(* IEC 61131-3 sources: SortJet_MasterSPS_Aufbau.fbsproj/11_MMI_Kommunikation, 12 files *)

(* ---- MMI_CONST.gvl ---- *)
(* METADATA
{
	"v3Meta": {
		"objectGuid": "b42c2871-ef06-40a1-9ac4-06faa3b26b72"
	}
}
*)
{attribute 'allow_unqualified_access'}
NAMESPACE MMI_CONST
VAR_GLOBAL CONSTANT

  sSpsVersion                                      : STRING(25) := 'ISO Sortierung V4.0.0.0';

// ************************ START SPS Nachrichtennummern *****************

  SB0_SPS_SPSVERSION                                 : WORD := 32768;
  SB0_SPS_MSG_ERROR                                  : WORD := 32767;
  SB0_SPS_ERROR                                      : WORD := 32766;
  SB0_SPS_WARNUNG                                    : WORD := 32765;
  SB0_SPS_HINWEIS                                    : WORD := 32764;
  SB0_SPS_PARAMETER_CRC                              : WORD := 32763;
  SB0_SPS_DEBUG                                      : WORD := 32762;
  SB0_SPS_DEBUG_TRACE                                : WORD := 32761; // Nachricht die in ein seperates Log-File geschrieben wird ( Void- Message )
  SB0_SPS_LOGSTRING                                  : WORD := 32770; // Nachricht um einen String (60 Zeichen) in das Log zu schreiben

// Nachricht von der SPS zum MMI
  SB0_SPS_SETBETRIEBSART                             : WORD :=  1;
  SB0_SPS_SORTIERUNGQUITTINPUTINQUEUE                : WORD :=  2;
  SB0_SPS_SORTIERUNGQUITTUNGVONISOLINIE              : WORD := 11;
  SB0_SPS_SORTIERUNGQUITTEXTRACTIONSHUTTLEDATA       : WORD := 13;
  SB0_SPS_SORTIERUNGRACKINPOS                        : WORD := 19;
  SB0_SPS_SORTIERUNGRACKSTATIONSTATUS                : WORD := 23;
  SB0_SPS_ERRORMSG                                   : WORD := 30;
  SB0_SPS_TRANSPORTSTATE                             : WORD := 35; // Antwort auf Eckübergabenstatus 0 = Rücktransport / 1 = Weitertransoport
  SB0_SPS_RACKONLOADINGSTATION                       : WORD := 37; // Fächerwagen auf Füllstation angedockt
  SB0_SPS_RACKLOGIN                                  : WORD := 38; // Fächerwagen auf Einschleusestation angedockt
  SB0_SPS_STATUSRACKSTATION                          : WORD := 39; // Antwort auf die Nachricht: SB0_SPS_STATUSRACKSTATION
  SB0_SPS_SETSTATUSLOADINGSTATIONS                   : WORD := 44; // Antwort auf REQUESTSTATUSLOADINGSTATIONS mit 1 = frei; 2 = belegt; 0 = ungültig
  SB0_SPS_SHEETREMOVEDAPPROVALWALL                   : WORD := 45;
  SB0_SPS_SHEETONINPUTTABLE                          : WORD := 46;
  SB0_SPS_RACKPOSITION                               : WORD := 48;
  SB0_SPS_TURNSTATIONPOSITION                        : WORD := 49;

  SB0_SPS_SYSTEMCHECKFINISHED                        : WORD := 51;
  SB0_SPS_SETSHEETSONSHUTTLE                         : WORD := 53;
  SB0_SPS_STATIONSTATUS                              : WORD := 62;
  SBO_SPS_STATIONSEVENT                              : word := 65;
  SB0_SPS_GETSTATIONSTATUS                           : WORD := 67; // BEKOMMEN: Einen Station-Status bekommen -> SystemCheck: Ein/ Austransport etc.
  SB0_SPS_SETSHEETSONSTATION                         : WORD := 68; // Nachricht an die Oberflaeche fuer die Glasmessung auf den Stationen
  SB0_SPS_SORTIERUNGSHUTTLEPOS                       : WORD := 69;
  SB0_SPS_SHUTTLEVORABPOSITIONIERUNGUPDATE           : WORD := 70;
  SB0_SPS_QUITTSHUTTLEVORABPOSITIONIERUNG            : WORD := 71;
  SB0_SPS_SHUTTLEVORABPOSITIONIERUNGABBRUCH          : WORD := 72;
  SB0_SPS_SHUTTLEVORABPOSITIONIERUNGREADY            : WORD := 73;
  SB0_SPS_TRANSFERSHUTTLEFEHLER                      : WORD := 75;
  SB0_SPS_FACHAUFNAHMEDATEN                          : WORD := 76;
  SB0_SPS_TRANSFERSHUTTLECHECK_ABGESCHLOSSEN         : WORD := 77;
  SB0_SPS_LIFTEDTRANSFERSHUTTLEPOSITION              : WORD := 78;
  SB0_SPS_SCHNITTSTELLENDATENFREMDANLAGE             : WORD := 79;

  SB0_SPS_POSITIONMEASUREDATA                        : WORD := 81; // Fächerwagensuche: Wort 0 = (int) SPS Nr Shuttle  / Wort 1+2 = (real) Position rechte (?) Kante der Folie[-1 für nicht gefunden]
  SB0_SPS_HANDFUNKTION_STATUS                        : WORD := 82; // Antwort auf SB0_MMI_SETHANDFUNKTION [22]
  SB0_SPS_SHUTTLEHANDFUNKTION_STATUS                 : WORD := 83; // Antwort auf SB0_MMI_SETSHUTTLEHANDFUNKTION [23]
  SB0_SPS_WATCHDOGTEST                               : WORD := 99;
  SB0_SPS_TRANSFERSHUTTLEBUFFERSLOTPOS               : WORD := 100;
  SB0_SPS_QUIT_SHEET_ORDER                           : WORD := 101;
  SB0_SPS_QUIT_CARRIER_POSITION                      : WORD := 102;
  SB0_SPS_STATION_UPDATE                             : WORD := 110;

// ************************ START MMI Nachrichtennummern *****************
  SB0_MMI_SPSVERSION                                 : WORD := 32768;
  SB0_MMI_GETBETRIEBSART                             : WORD :=  1;
  SB0_MMI_SORTIERUNGINPUTINQUEUE                     : WORD :=  2;
  SB0_MMI_SORTIERUNGCHECKINPUTQUEUE                  : WORD :=  5;
  SB0_MMI_SORTIERUNGCANCELQUEUEDATA                  : WORD :=  7;
  SB0_MMI_SORTIERUNGCANCELISOLINEEVENT               : WORD :=  8; // ISO- Line Event stoppen [Cancel]
  SB0_MMI_SORTIERUNGCANCELSHUTTLEDATA                : WORD :=  9;
  SB0_MMI_SORTIERUNGFAECHERWAGENBALDVOLL             : WORD := 10; // Faecherwagen in der Station bald voll
  SB0_MMI_SORTIERUNGAUTOMATIKSTART                   : WORD := 11;
  SB0_MMI_SORTIERUNGAUTOMATIK_STOP                   : WORD := 12;
  SB0_MMI_SORTIERUNGINSERTEXTRACTIONSHUTTLEDATA      : WORD := 14;
  SB0_MMI_SORTIERUNGFAECHERWAGENWECHSEL              : WORD := 15;
  SB0_MMI_SETHANDFUNKTION                            : WORD := 22;
  SB0_MMI_SETSHUTTLEHANDFUNKTION                     : WORD := 23;
  SB0_MMI_MEASSURERESULT                             : WORD := 30; // Scheibenmessung OK -> Freigabe für die Eckübergabe des Sortjets  0 = nicht OK / 1 = OK
  SB0_MMI_ISOQUITTUNG                                : WORD := 31; // unabhängige Quittung der Sondergläser durch Tasterdruck anfordern
  SB0_MMI_RELEASERACKLOGIN                           : WORD := 39; // Freigabe, dass der Fächerwagen eingeschleußt werden darf
  SB0_MMI_GETSTATUSRACKSTATION                       : WORD := 40; // Anfrage vom MMI nach dem Status einer EINZELNEN Fächerwagenstation => belegt, Muting OK, RFID-Nr.
  SB0_MMI_DOCKRACK                                   : WORD := 41; // Freigabe den AGV Fächerwagen einzuschleusen bzw. das Tor zu öffnen  /  release to open the door for the AGV harp rack
  SB0_MMI_REQUESTSTATUSLOADINGSTATIONS               : WORD := 43; // Anfrage der Oberfläche welche Fächerwagenbeladestationen belegt sind
  SB0_MMI_SETSLOTSFORSHUTTLECHECK                    : WORD := 44; // Anfrage der aktuellen Shuttlepositionnen für den bevorstehenden Check der Maschine
  SB0_MMI_REQUESTTILTSTATION                         : WORD := 51;
  SB0_MMI_SHUTTLEVORABPOSITIONIERUNG                 : WORD := 53; // Shuttle Vorapositionieren falls ein Transfershuttle (welches benötigt wird) gerade beschäftigt ist
  SB0_MMI_FACHAUFNAHMESTART                          : WORD := 55;
  SB0_MMI_POSITIONMEASUREONOFF                       : WORD := 56; // FächerwagenSUCHE    Wort 0 = (int) 1 für AN oder 0 für AUS / Wort 2 = (int) SPS Nr Shuttle
  SB0_MMI_STATIONSTATUS                              : WORD := 67; // Stationsstatus [Antwort in welchem Modus sich die Station befunden hat -> SystemCheck]
  SB0_MMI_SYSTEMCHECKSTATION                         : WORD := 68; // Stationsstatus [Antwort in welchem Modus sich die Station befunden hat -> SystemCheck]
  SB0_MMI_GETSORTIERUNGSHUTTLEPOS                    : WORD := 69;
  SB0_MMI_IOANZEIGE_AKTIVIEREN_DEAKTIVIEREN          : WORD := 70; // Anzeige der IO´s im MMI Service  WORT 0: 1 = sichtbar / 0 = unsichtbar
  SB0_MMI_AUFTRAGSDATEN_FREMDANLAGE                  : WORD := 71; // Uebertragen von Daten ueber eine Hardwareschnittstelle \ DPD-Koppler an eine Fremdanlage
  SB0_MMI_SHUTTLE_INFORMATION                        : WORD := 72; // Uebertragen von Daten waehrend der Shuttle-Positionierung
  SB0_MMI_TRANSFERSHUTTLECHECK                       : WORD := 76; // Hinweis: Systemcheck mit Transfershuttles da Glas aus dem Speicher raus stand
  SB0_MMI_LIFTTRANSFERSHUTTLE                        : WORD := 77;
  SB0_MMI_DURCHTRANSPORT                             : WORD := 80;
  SB0_MMI_RESET_ETHERCAT                             : WORD := 81;
  SB0_MMI_WATCHDOGTEST                               : WORD := 99;
  SB0_MMI_TRANSFERSHUTTLEBUFFERSLOTCHECK             : WORD := 100;
  SB0_MMI_SHEET_ORDER                                : WORD := 101;
  SB0_MMI_DRIVEOVERRIDE                              : WORD := 102;
  SB0_MMI_START_BELT_CLEANING                        : WORD := 103;
  SB0_MMI_CARRIER_POSITIONING                        : WORD := 104;
  SB0_MMI_TS_REPOSITIONING_LITES                     : WORD := 110;

END_VAR

END_NAMESPACE

(* ---- MMI_Vars.gvl ---- *)
(* METADATA
{
	"v3Meta": {
		"objectGuid": "3eb4075d-cf2f-4b71-9fd2-f0699e9e6b81"
	}
}
*)
{attribute 'allow_unqualified_access'}
NAMESPACE MMI_Vars
VAR_GLOBAL
  bgMMIOK : BOOL;

  // SPS -> MMI
  dwSps2MmiHandfunktionenStatus                   : DWORD;
  wSps2MmiErrorShuttleNumber                      : WORD;
  wSps2MmiErrorShuttleSchritt                     : WORD;
  wSps2MmiErrorNumber                             : WORD;
  wSps2FaecherwagenStart                          : WORD;
  wSps2MmiStatusforStation                        : WORD; // Anfrage der Eckübergabe (Nr) wohin die Einlaufende Scheibe soll

  wSps2MmiQuittISOLineNr                          : WORD;
  wSPS2MMIStationsNummer                          : WORD;
  wSPS2MMITRANSPORTSTATE                          : WORD;
  wSPS2MMITransportstateStation                   : WORD;
  rSPS2MMITransportStateLenght                    : REAL;
  rSPS2MMITransportStateHigh                      : REAL;
  wSPS2MMITransportstateGap                       : WORD;
  wSps2FaecherwagenStationNr                      : WORD;
  wSps2MmiInputtableNummer                        : WORD;
  wSps2MmiRackNumber                              : WORD;

  wSps2MmiWatchDogTestCount                       : WORD;

  // SB0_SPS_GLAS_SOLLPOSITION_ERREICHT
  wgSps2MmiShuttleNr                              : WORD;
  wSps2MmiRackPositionNummer                      : WORD;
  wSps2MmiRackPosition                            : WORD;
  wSps2MmiRackStatus                              : WORD;
  wgSps2MmiPosDrehStation                         : WORD;
  wgSps2MmiOldPosDrehStation                      : WORD;
  wgSps2MmiDrehStation                            : WORD;
  wSps2MmiCheckArea                               : WORD;
  wSps2MmiCheckSuccessful                         : WORD;
  wSps2MmiMeasureShuttleNummer                    : WORD;
  wSps2MmiErrorShuttlePosition4                   : WORD;
  wSps2MmiErrorShuttlePosition5                   : WORD;
  wSps2MmiErrorShuttlePosition6                   : WORD;
  wSps2MmiErrorShuttlePosition7                   : WORD;
  wSps2MmiErrorShuttlePosition8                   : WORD;
  wSps2MmiErrorShuttlePosition9                   : WORD;

  // Debug
  wSps2MmiDebugLogWord1                           : WORD;
  wSps2MmiDebugLogWord2                           : WORD;
  wSps2MmiDebugLogWord3                           : WORD;
  wSps2MmiDebugLogWord4                           : WORD;
  wSps2MmiDebugLogWord5                           : WORD;
  wSps2MmiDebugLogWord6                           : WORD;
  wSps2MmiDebugLogWord7                           : WORD;
  wSps2MmiDebugLogWord8                           : WORD;
  wSps2MmiDebugLogWord9                           : WORD;

  // SB0_SPS_STATIONEVENT
  wSPS2MMIStationEventStatus                      : WORD;

  // SB0_SPS_QUIT_SHEET_ORDER
  wSps2MmiZielStation                             : WORD;
  wSps2MmiQuellStation                            : WORD;
  wSps2MmiZielWand                                : WORD;
  wSps2MmiQuellWand                               : WORD;
  wSPS2MMIAuftragstyp                             : WORD;
  dwSPS2MMIGenutzteSauger                         : DWORD;

  // Offset
  // Nachricht: SB0_SPS_STATUSISOLINIE
  wSPS2MMIISOLinieNummer                          : WORD;
  wSPS2MMIShuttleNummer                           : WORD;
  wSPS2MMIShuttleKippenStatus                     : WORD;
  // SB0_SPS_LIFTEDTRANSFERSHUTTLEPOSITION
  wSps2MmiValidierungsPosition                    : REAL;
  wSps2MmiValidierungsSpeicher                    : WORD;
  wSps2MmiValidierungsFach                        : WORD;

  // SB0_SPS_TRANSFERSHUTTLEFEHLER
  wSps2MmiFehlertyp                               : WORD;

  // SB0_SPS_TRANSFERSHUTTLECHECK_ABGESCHLOSSEN
  wSps2MmiValidierungsStatus                      : WORD;

  // SB0_SPS_SORTIERUNGQUITTEXTRACTIONSHUTTLEDATA
  wSps2MmiQuittierungVortransportStationsNr1      : WORD;
  wSps2MmiQuittierungVortransportStationsNr2      : WORD;
  wSps2MmiQuittierungVortransportStatus           : WORD;
  rSps2MmiQuittierungVortransportWegStrecke       : REAL;

  // Stationsstatus
  wSPS2MMIStationsStatusWord1                     : WORD;
  wSPS2MMIStationsStatusWord2                     : WORD;

 // SB0_SPS_SETSHEETSONSTATION
  rSps2MmiMessungScheibenlaenge                   : REAL;
  wSps2MmiMessungStationNummer                    : WORD;
  wSps2MmiMessungSlotNummer                       : WORD;
  iSps2MmiMessungScheibenanzahl                   : INT;

 // Fachaufnahme
  wSPS2MMIFachaufnahmeAnalogwert                  : WORD;
  rSPS2MMIFachaufnahmePosition                    : REAL;

  // Nachricht: SB0_SPS_SETSTATUSLOADINGSTATIONS
  awSps2MmiStatusFaecherwagenstationen             : ARRAY [0..29] OF WORD;

  // Verfahrlogik_Neu
  wSps2MmiQuittVorabShuttleNr                     : WORD;
  rgSPS2MMIExtractionShuttlePosition              : REAL;
  rgSPS2MMIExtractionShuttlePositionHub           : REAL;
  rSps2MmiShuttlePosition                         : ARRAY [0..30] OF REAL; // Liste fuer SB0_SPS_SORTIERUNGSHUTTLEPOS [SendShuttlePosition]
  rSps2MmiPosition                                : REAL;  // Position fuer Einzelnachrichten [VORABPOSITIONIERUNG ABBRUCH/READY, POSITIONMEASUREDATA]
  wSps2ShuttleStopped                             : ARRAY [cERSTES_SHUTTLE..cLETZTE_STATION] OF WORD;

  rgSPS2MMIExtractionShuttleGefahrenerWeg         : REAL;
  rSps2MmiMeasureResult                           : ARRAY [0..10] OF REAL;

  dwSps2MmiWartezeit                              : DWORD; // ZEIT-WERT MMI-STATISTIK: Beschreibt die Zeit zwischen Anlegeauftrag und dem betaetigen des Tasters zum Eintransport

  // SB0_SPS_STATUSRACKSTATION
  igRackStationNumber                             : INT;   // Fächerwagenstationsnummer / Harp Rack Station
  wgRackPresent                                   : WORD;  // BOOL (0 oder 1)
  igRackNumber                                    : INT;   // RFID Number
  wgWriteSuccess                                  : WORD;  // Zeigt an wie das Schreiben des RFID-Chips verlaufen ist (0=none|1=success|2=error)

  wSps2Mmi_CarrierStation                         : WORD;
  wSps2Mmi_CarrierPosition                        : REAL;

  wSps2Mmi_SationsNummer                          : WORD;
  wSps2Mmi_NachrichtenIndex                       : WORD;
  wSps2Mmi_NachrichtenAnzahl                      : WORD;
  wSps2Mmi_AnzahlScheiben                         : WORD;
  adwSps2Mmi_Daten_1                              : ARRAY [0..3] OF DWORD;
  adwSps2Mmi_Daten_2                              : ARRAY [0..3] OF DWORD;
  adwSps2Mmi_Daten_3                              : ARRAY [0..3] OF DWORD;

  wSps2MmiKorrekturStatus                         : WORD;

  stStationUpdate                                  : StationUpdate_ST;

  // ---------------------------------------------------------------------------------------
  // MERKER - NACHRICHTEN
  //
  // Hinweis:
  // - Trigger das ein Auftrag in der SPS zugewiesen und bearbeitet wird
  // ---------------------------------------------------------------------------------------

  M_SB0_MMI_SortierungInputInQueue                : BOOL;
  M_SB0_MMI_SortierungCheckInputQueue             : BOOL;
  M_SB0_MMI_SORTIERUNGCANCELISOLINEEVENT          : BOOL; // Intern: ISO- Linie Event abbrechen [CANCEL]

  M_SB0_MMI_SortierungInsertExtractionShuttleData : BOOL;// NEU
  M_SB0_MMI_TS_REPOSITIONING_LITES                : BOOL;
  M_SB0_MMI_SortierungFaecherwagenwechsel         : BOOL;
  M_SB0_MMI_SORTIERUNGFAECHERWAGENBALDVOLL        : BOOL;
  M_SB0_MMI_SortierungCancelShuttleData           : BOOL;
  M_SB0_MMI_SORTIERUNGCANCELQUEUEDATA             : BOOL;
  M_SB0_MMI_SortierungAutomatik_Stop              : BOOL;
  M_SB0_MMI_SORTIERUNGAUTOMATIKSTART              : BOOL;
  M_SB0_MMI_SYSTEMCHECKSTATION                    : BOOL;
  M_SB0_MMI_STATIONSTATUS                         : BOOL;
  M_SB0_MMI_MEASSURERESULT                        : BOOL;
  M_SB0_MMI_ISOQUITTUNG                           : BOOL;
  M_SB0_MMI_GETSTATUSRACKSTATION                  : BOOL;
  M_SB0_MMI_REQUESTSTATUSLOADINGSTATIONS          : BOOL;
  M_SB0_MMI_REQUESTTILTSTATION                    : BOOL;
  M_SB0_MMI_GETSORTIERUNGSHUTTLEPOS               : BOOL; // VERFAHRLOGIK
  M_SB0_MMI_SHUTTLEVORABPOSITIONIERUNG            : BOOL; // VERFAHRLOGIK
  M_SB0_MMI_SHEET_ORDER_SHUTTLE                   : BOOL;
  M_SB0_MMI_SHEET_ORDER_STATION                   : BOOL;
  M_SB0_MMI_RELEASERACKLOGIN                      : BOOL;
  M_SB0_MMI_DOCKRACK                              : BOOL;
  M_SB0_MMI_CARRIER_POSITIONING                   : BOOL;
  M_SB0_MMI_DRIVEOVERRIDE                         : BOOL;
  M_SB0_MMI_WATCHDOGTEST                          : BOOL;
  M_SB0_MMI_RESET_ETHERCAT                        : BOOL;
  M_SB0_MMI_IOANZEIGE_AKTIVIEREN_DEAKTIVIEREN     : BOOL; // IOs Anzeigen

  M_SB0_MMI_AUFTRAGSDATEN_FREMDANLAGE             : BOOL; // MERKER: Auftragsdaten fuer die Fremdanlage

  M_SB0_MMI_SHUTTLE_INFORMATION                   : BOOL; // MERKER: Shuttledaten- Waehrend einer Verfahrbewegung senden

  M_SB0_MMI_POSITIONMEASUREONOFF                  : BOOL;
  M_SB0_MMI_TRANSFERSHUTTLECHECK                  : BOOL; // Merker: Systemcheck mit Transfershuttles da Glas aus dem Speicher raus stand

  M_SB0_MMI_ANFORDERUNG_PUFFER_AUSFAHREN          : BOOL;
  M_SB0_MMI_ANFORDERUNG_PUFFER_EINFAHREN          : BOOL;

// ------------------------------------------

 M_Send_MaschineStatus : BOOL;
  // ----- Sps Message Queue -----
 smqSpsMessageQueue : SpsMessageQueue;

// MMI -> SPS
 tMmi2SpsInfo : Mmi2SpsInfo;

// Fehlerparameter zur Übergabe ans MMI
 wpgFehlerdaten : ARRAY[0..25] OF WORD;

// SPS -> MMI
 awSPS2MMIMaschineStatusWord : ARRAY[1..12] OF WORD;

END_VAR

END_NAMESPACE

(* ---- TCP_Global.gvl ---- *)
(* METADATA
{
	"v3Meta": {
		"objectGuid": "822ea3bc-9f3a-414f-ba8a-dc2da6267ba8"
	}
}
*)
{attribute 'allow_unqualified_access'}
NAMESPACE TCP_Global
VAR_GLOBAL
  g_bCallbackRegistered : BOOL;
  bgTcpConnected        : BOOL;
  bgCallback_ONLINE_CHANGE : BOOL;
  bgCallback_BEFORE_RESET : BOOL;
  bgCallback_BEFORE_DOWNLOAD : BOOL;
  bgCallback_Shutdown : BOOL;
  bgSteuerung_Eckelmann : BOOL := TRUE;
END_VAR
VAR_GLOBAL CONSTANT
  // Nachrichtenkonstanten der TCP Schnitstelle
  cMsg_Watchdog      : WORD := 16#0001;
  cMsg_MsgBlock      : WORD := 16#0002;
  cMsg_ControlSystem : WORD := 16#0003;
  cMsg_IOSystem      : WORD := 16#0004;
  cMsg_Drives        : WORD := 16#0005;
  cMsg_MsgDirect     : WORD := 16#0006;
  cMsg_MsgDirectAck  : WORD := 16#0007;
END_VAR
END_NAMESPACE

(* ---- MsgInterpret.fn.st ---- *)
(* METADATA
{
	"v3Meta": {
		"objectGuid": "c5198d31-be99-460b-8031-114f442e3133"
	}
}
*)
FUNCTION MsgInterpret : BOOL
VAR_INPUT
  tSpsMessage : SpsMessage;
END_VAR
VAR
  wlIndex : WORD;
  wlTemp  : WORD;
END_VAR

CASE( tSpsMessage.wAuftrag )OF

  // MSG 1
  // Anfrage des Maschinenstatuses
  SB0_MMI_GETBETRIEBSART:
    M_Send_MaschineStatus := TRUE;

  // MSG 2
  // Auftrag für den Anlegetisch (Start_Station)
  SB0_MMI_SortierungInputInQueue:
    tMmi2SpsInfo.wSortierungsInQueueLineNr         := HMI_GetWORD(ADR(tSpsMessage.awDaten[0]));  // Liniennr. wo das Glas aufgelegt werden soll
    tMmi2SpsInfo.wSortierungsInputInQueueStationNr := HMI_GetWORD(ADR(tSpsMessage.awDaten[1])); // Tischnummer des Anlegetisches
    tMmi2SpsInfo.rInputInQueueLaenge               := HMI_GetREAL(ADR(tSpsMessage.awDaten[2]));
    tMmi2SpsInfo.rInputInQueueHoehe                := HMI_GetREAL(ADR(tSpsMessage.awDaten[4]));
    tMmi2SpsInfo.rInputInQueueDicke                := HMI_GetREAL(ADR(tSpsMessage.awDaten[6]));
    tMmi2SpsInfo.wInsertInputShuttleDataCoatedSide := HMI_GetWORD(ADR(tSpsMessage.awDaten[8]));// Coated_Side
    tMmi2Spsinfo.wSortierungInQueueSheetOut        := HMI_GetWORD(ADR(tSpsMessage.awDaten[9]));  // 0=Glas für Sortjet; 1= Glas nicht für Sortjet

    tMmi2SpsInfo.wModellStatus         := HMI_GetWORD(ADR(tSpsMessage.awDaten[11]));
    tMmi2SpsInfo.rModellVersatzVorne   := HMI_GetREAL(ADR(tSpsMessage.awDaten[12]));
    tMmi2SpsInfo.rModellversatzHinten  := HMI_GetREAL(ADR(tSpsMessage.awDaten[14]));
    tMmi2SpsInfo.rModellVersatzVorne2  := HMI_GetREAL(ADR(tSpsMessage.awDaten[16]));
    tMmi2SpsInfo.rModellversatzHinten2 := HMI_GetREAL(ADR(tSpsMessage.awDaten[18]));
    tMmi2SpsInfo.wPrintStatus          := HMI_GetWORD(ADR(tSpsMessage.awDaten[20]));
    tMmi2SpsInfo.wSourceTable          := HMI_GetWORD(ADR(tSpsMessage.awDaten[21]));
    tMmi2SpsInfo.wSlotZielStation      := HMI_GetWORD(ADR(tSpsMessage.awDaten[22]));

    M_SB0_MMI_SortierungInputInQueue := TRUE;

  // MSG 5
  // Starten des SystemCheck
  SB0_MMI_SortierungCheckInputQueue:
    tMmi2SpsInfo.wCheckArea      := HMI_GetWORD(ADR(tSpsMessage.awDaten[0]));
    tMmi2SpsInfo.wCheckRelease   := HMI_GetWORD(ADR(tSpsMessage.awDaten[1]));
    M_SB0_MMI_SortierungCheckInputQueue := TRUE;

  // MSG 7
  // Beliebige Station irgendeiner Linie die Daten löschen
  SB0_MMI_SORTIERUNGCANCELQUEUEDATA:   // SB0_MMI_SortierungDelete:
    tMmi2SpsInfo.wDeleteStationNr   := HMI_GetWORD(ADR(tSpsMessage.awDaten[0])); // Tischnummer des Anlegetisches
    tMmi2SpsInfo.wDeleteStationSlot := HMI_GetWORD(ADR(tSpsMessage.awDaten[1])); // Wandnummer  des Anlegetisches
    M_SB0_MMI_SORTIERUNGCANCELQUEUEDATA := TRUE;

  // MSG 8
  // Abbruch des offenen ISO Line Events
  SB0_MMI_SORTIERUNGCANCELISOLINEEVENT:
    M_SB0_MMI_SORTIERUNGCANCELISOLINEEVENT := TRUE;

  // MSG 9
  // Auftrag des entsprechenden Shuttles löschen
  SB0_MMI_SortierungCancelShuttleData:
    tMmi2SpsInfo.wCancelShuttleDataShuttleNr := HMI_GetWORD(ADR(tSpsMessage.awDaten[0]));
    M_SB0_MMI_SortierungCancelShuttleData := TRUE;

  // MSG 11
  // Start Automatik Foerder Transport der Glastransportstationen
  SB0_MMI_SORTIERUNGAUTOMATIKSTART:
    tMmi2SpsInfo.wAutomatikStartTransportLineNr := HMI_GetWORD(ADR(tSpsMessage.awDaten[0]));
    M_SB0_MMI_SORTIERUNGAUTOMATIKSTART := TRUE;

  // MSG 12
  (* Hinweis:
     - Nachricht von der Oberflaeche das ein Automatikkreis gestopt werden soll / muss
       => Index[0] Angabe welcher Automatikkreis gestoppt werden soll
       => Index[1] Angabe welche Automatikkreise schon gestoppt sind
     - Falls schon einer der beiden Kreise gestoppt wurde, steht im 2. Datenwort eine 3.
       Wenn eine 3 vorkommt, dann diese übernehmen um beide Autokreise, inkl. den Transfershuttlen stoppen
  *)
  SB0_MMI_SortierungAutomatik_Stop:
    tMmi2SpsInfo.wAutomatikStopArea     := HMI_GetWORD(ADR(tSpsMessage.awDaten[0]));
    tMmi2SpsInfo.wAutomatikStoppedAreas := HMI_GetWORD(ADR(tSpsMessage.awDaten[1]));
    M_SB0_MMI_SortierungAutomatik_Stop := TRUE;

  // MSG 14
  // Vorpositionier der Scheiben im Speicher (Transfershuttle)
  SB0_MMI_SortierungInsertExtractionShuttleData:
    tMmi2SpsInfo.wVortransportNummer_TS1       := HMI_GetWORD(ADR(tSpsMessage.awDaten[0]));
    tMmi2SpsInfo.rVortransportSollPosition_TS1 := HMI_GetREAL(ADR(tSpsMessage.awDaten[1]));
    tMmi2SpsInfo.rVortransportStrecke          := HMI_GetREAL(ADR(tSpsMessage.awDaten[3]));
    tMmi2SpsInfo.wVortransportNummer_TS2       := HMI_GetWORD(ADR(tSpsMessage.awDaten[5]));
    tMmi2SpsInfo.rVortransportSollPosition_TS2 := HMI_GetREAL(ADR(tSpsMessage.awDaten[6]));
    tMmi2SpsInfo.wSlotThickness                := HMI_GetWORD(ADR(tSpsMessage.awDaten[8])); // 0-thin;1-thick

    M_SB0_MMI_SortierungInsertExtractionShuttleData := TRUE;

  // MSG 10
  // Faecherwagen in der Station bald voll: Anzeige an der Station
  SB0_MMI_SORTIERUNGFAECHERWAGENBALDVOLL:
    tMmi2SpsInfo.wSps2FaecherwagenStationNr  := HMI_GetWORD(ADR(tSpsMessage.awDaten[0]));   // Stationsnummer
    M_SB0_MMI_SORTIERUNGFAECHERWAGENBALDVOLL := TRUE;

  // MSG 15
  // Fächerwagenwechsel auch von verschiedenen Stationen möglich
  SB0_MMI_SORTIERUNGFAECHERWAGENWECHSEL:
    tMmi2SpsInfo.wFaecherwagenwechsel       := HMI_GetWORD(ADR(tSpsMessage.awDaten[0]));   // DestStation / Zielstation
    tMmi2SpsInfo.wSps2FaecherwagenStationNr := HMI_GetWORD(ADR(tSpsMessage.awDaten[1]));   // SourceStation / Startstation
    M_SB0_MMI_SortierungFaecherwagenwechsel:=TRUE;

  // MSG 22
  // HANDFUNKTIONEN: Stationen
  SB0_MMI_SetHandfunktion:
    FOR wlIndex := 0 TO (tSpsMessage.wLaenge-1) BY 6 DO

      IF ( HMI_GetWORD(ADR(tSpsMessage.awDaten[0])) >= cERSTE_FAECHERWAGENSTATIONS_NR ) THEN
        adwgHandfunktionenFaecherwagenStationen[HMI_GetWORD(ADR(tSpsMessage.awDaten[wlIndex/2]))] := HMI_GetDWORD(ADR(tSpsMessage.awDaten[( (wlIndex)/2 )+1]));
      ELSE
        adwgHandfunktionenStationen[HMI_GetWORD(ADR(tSpsMessage.awDaten[wlIndex/2]))] := HMI_GetDWORD(ADR(tSpsMessage.awDaten[( (wlIndex)/2 )+1]));
      END_IF

    END_FOR

  // MSG 23
  // HANDFUNKTIONEN: Shuttle
  SB0_MMI_SetShuttleHandFunktion:
    IF HMI_GetWORD(ADR(tSpsMessage.awDaten[0])) >= cERSTE_STATION THEN
      FOR wlIndex := 0 TO (tSpsMessage.wLaenge-1) BY 6 DO
        adwgHandfunktionenStationen[HMI_GetWORD(ADR(tSpsMessage.awDaten[wlIndex/2]))] := HMI_GetDWORD(ADR(tSpsMessage.awDaten[( (wlIndex)/2 )+1]));
      END_FOR
    ELSIF HMI_GetWORD(ADR(tSpsMessage.awDaten[0])) >= cERSTES_TRANSFERSHUTTLE THEN
      FOR wlIndex := 0 TO (tSpsMessage.wLaenge-1) BY 6 DO
        adwgHandfunktionenTransfershuttle[HMI_GetWORD(ADR(tSpsMessage.awDaten[wlIndex/2]))] := HMI_GetDWORD(ADR(tSpsMessage.awDaten[( (wlIndex)/2 )+1]));
      END_FOR
    ELSE
      FOR wlIndex := 0 TO (tSpsMessage.wLaenge-1) BY 6 DO
        adwgHandfunktionenShuttle[HMI_GetWORD(ADR(tSpsMessage.awDaten[wlIndex/2]))] := HMI_GetDWORD(ADR(tSpsMessage.awDaten[( (wlIndex)/2 )+1]));
      END_FOR
    END_IF

  // MSG 30
  // Scheibenmessung OK -> Freigabe für die Eckübergabe des Sortjets  0 = nicht OK / 1 = OK
  SB0_MMI_MEASSURERESULT:
    M_SB0_MMI_MEASSURERESULT:=TRUE;
    tMmi2SpsInfo.wFreigabe               := HMI_GetWORD(ADR(tSpsMessage.awDaten[0]));// Freigabe
    tMmi2SpsInfo.wMmiNummerAnlegeStation := HMI_GetWORD(ADR(tSpsMessage.awDaten[1]));

  // MSG 31
  // Unabhaengige Quittung der Sondergläser durch Tasterdruck anfordern
  SB0_MMI_ISOQUITTUNG:
    M_SB0_MMI_ISOQUITTUNG:=TRUE;
    tMmi2SpsInfo.wISOStation    := HMI_GetWORD(ADR(tSpsMessage.awDaten[0])); (* Tischnummer des Anlegetisches *)// Liniennummer
    tMmi2SpsInfo.wISOAuftragsID := HMI_GetWORD(ADR(tSpsMessage.awDaten[1]));// Auftrags ID

  // MSG 39
  // Bestaetigung der Faecherwagenanmeldung vom MMI
  SB0_MMI_RELEASERACKLOGIN:
    M_SB0_MMI_RELEASERACKLOGIN := TRUE;
    tMmi2SpsInfo.wSps2FaecherwagenStationNr  := HMI_GetWORD(ADR(tSpsMessage.awDaten[0])); // Stationsnummer wo der Wagen eingeschleust werden soll
    tMmi2SpsInfo.wlFreigabeEinschleuseJaNein := HMI_GetWORD(ADR(tSpsMessage.awDaten[1])); // Freigabe zum Einschleusen = 1 / Freigegebenen Wagen wieder löschen = 0

  // MSG 40
  // Anfrage vom MMI nach dem Status einer EINZELNEN Fächerwagenstation => belegt, Muting OK, RFID-Nr.
  SB0_MMI_GETSTATUSRACKSTATION:
    M_SB0_MMI_GETSTATUSRACKSTATION := TRUE;
    tMmi2SpsInfo.wSps2FaecherwagenStationNr := HMI_GetWORD(ADR(tSpsMessage.awDaten[0])); // Stationsnummer wo angefragt wird
  // - Freigabe eines mittles AGV eingeschleusten Wagen das Tor zu öffnen

  // MSG 41
  SB0_MMI_DOCKRACK:
    M_SB0_MMI_DOCKRACK := TRUE;
    tMmi2SpsInfo.wSps2FaecherwagenStationNr := HMI_GetWORD(ADR(tSpsMessage.awDaten[0]));

  // MSG 43
  (* Hinweis [FAECHERWAGEN]:
     - MMI Anfrage, welche Fächerwagenstationen belegt sind
       => <igIndexFaecherwagenDaten> wird zum Auslesen der Daten benoetigt da hier der Index bei "0" anfaengt
  *)
  SB0_MMI_REQUESTSTATUSLOADINGSTATIONS:
    igIndexFaecherwagenDatenEmpfangen := 0;
    FOR wlIndex := cERSTE_FAECHERWAGENSTATIONS_NR TO cLETZTE_FAECHERWAGENSTATIONS_NR DO
      tMmi2SpsInfo.awAnfrageStatusDerFaecherwagenstation[wlIndex] := HMI_GetWORD(ADR(tSpsMessage.awDaten[igIndexFaecherwagenDatenEmpfangen]));
      igIndexFaecherwagenDatenEmpfangen := igIndexFaecherwagenDatenEmpfangen + 1;
    END_FOR
    M_SB0_MMI_REQUESTSTATUSLOADINGSTATIONS := bgEtherCatOK;

  // MSG 51
  SB0_MMI_REQUESTTILTSTATION:
    tMmi2SpsInfo.wSortierungsInputSwingStationNr := HMI_GetWORD(ADR(tSpsMessage.awDaten[0])); // Stationsnummer
    M_SB0_MMI_REQUESTTILTSTATION := TRUE;

  // MSG 53
  // Positionierung ueber die Oberflaeche [Verfahrlogik]
  SB0_MMI_SHUTTLEVORABPOSITIONIERUNG:
    tMmi2SpsInfo.wVorabStationsNr        := HMI_GetWORD(ADR(tSpsMessage.awDaten[0]));
    tMmi2SpsInfo.rVorabPositionierung    := HMI_GetREAL(ADR(tSpsMessage.awDaten[1]));
    tMmi2SpsInfo.rVorabUpdateZeit        := HMI_GetREAL(ADR(tSpsMessage.awDaten[3]));
    tMmi2SpsInfo.wVorabAuftragstyp       := HMI_GetWORD(ADR(tSpsMessage.awDaten[16]));
    M_SB0_MMI_SHUTTLEVORABPOSITIONIERUNG := TRUE;

  // MSG 55
  // Fachaufnahme
  SB0_MMI_FACHAUFNAHMESTART:
    wlTemp := HMI_GetWORD(ADR(tSpsMessage.awDaten[0]));
    AutomatischeFachaufnahme.bpStarteFachaufnahme := wlTemp.0;
    AutomatischeFachaufnahme.wpMMINummer          := HMI_GetWORD(ADR(tSpsMessage.awDaten[2]));

  // MSG 56
  // Shuttle Fächerwagen ausmessen
  SB0_MMI_POSITIONMEASUREONOFF:
    tMmi2SpsInfo.wShuttleNummerFWSuche := HMI_GetWORD(ADR(tSpsMessage.awDaten[0]));
    tMmi2SpsInfo.wShuttleFWSucheAN_AUS := HMI_GetWORD(ADR(tSpsMessage.awDaten[1]));

    M_SB0_MMI_POSITIONMEASUREONOFF := TRUE;

  // MSG 67
  // STATUS: Stationen (SystemCheck)
  SB0_MMI_STATIONSTATUS:
    tMmi2SpsInfo.wStationsNummer      := HMI_GetWORD(ADR(tSpsMessage.awDaten[0])); // Station Nr.
    tMmi2SpsInfo.wStationsStatusWord1 := HMI_GetWORD(ADR(tSpsMessage.awDaten[1])); // Manueller Modus
    tMmi2SpsInfo.wStationsStatusWord2 := HMI_GetWORD(ADR(tSpsMessage.awDaten[2])); // Schleifen
    tMmi2SpsInfo.wStationsStatusWord3 := HMI_GetWORD(ADR(tSpsMessage.awDaten[3])); // Modelle
    tMmi2SpsInfo.wStationsStatusWord4 := HMI_GetWORD(ADR(tSpsMessage.awDaten[4])); // Ebene /Slotnummer
    tMmi2SpsInfo.wStationsStatusWord5 := HMI_GetWORD(ADR(tSpsMessage.awDaten[5])); // Drehposition
    tMmi2SpsInfo.wStationsStatusWord6 := HMI_GetWORD(ADR(tSpsMessage.awDaten[6])); // Blockiert
    tMmi2SpsInfo.wStationsStatusWord7 := HMI_GetWORD(ADR(tSpsMessage.awDaten[7])); // 0 = inaktiv | 1 = aktiv

    M_SB0_MMI_STATIONSTATUS := TRUE;

  // MSG 68
  // DATEN FÜR DEN SYSTEMCHECK
  SB0_MMI_SYSTEMCHECKSTATION:
    M_SB0_MMI_SYSTEMCHECKSTATION := TRUE;
    tMmi2SpsInfo.wSystemCheckStationMmiNummer          := HMI_GetWORD(ADR(tSpsMessage.awDaten[0])); // Stationsnummer
    tMmi2SpsInfo.wSystemCheckStationScheibenanzahl     := HMI_GetWORD(ADR(tSpsMessage.awDaten[1])); // Scheibenanzahl [Gibt an wieviele Scheiben auf der Station sind]
    tMmi2SpsInfo.wSystemCheckStationZielstation        := HMI_GetWORD(ADR(tSpsMessage.awDaten[2])); // Zielstation (lt. MMI)
    tMmi2SpsInfo.wSystemCheckStationLetzteScheibe      := HMI_GetWORD(ADR(tSpsMessage.awDaten[3])); // Die Station ist bei gesetztem Bit- voll beladen
    tMmi2SpsInfo.wSystemCheckStationBeschichtungsSeite := HMI_GetWORD(ADR(tSpsMessage.awDaten[4])); // Beschichtungsseite
    tMmi2SpsInfo.wSystemCheckStationTyp                := HMI_GetWORD(ADR(tSpsMessage.awDaten[5])); // Hinweis: Kann benutzt werden fuer spezielle Bedingungen -> TeutoGlas Ausrichttypen fuer die Station 211 [Ausrichtfoerderer]
    tMmi2SpsInfo.wSystemCheckStationSlot               := HMI_GetWORD(ADR(tSpsMessage.awDaten[6])); // Wandnr
    tMmi2SpsInfo.rSystemCheckStationSollPosition       := HMI_GetREAL(ADR(tSpsMessage.awDaten[7])); // Hinweis: Gibt Auskunft ueber die Position an der z.B. ein Antrieb gestanden hat / stehen soll
    tMmi2SpsInfo.rSystemCheckStationScheibenlaenge     := HMI_GetREAL(ADR(tSpsMessage.awDaten[9])); // ** NEU Startposition als ABS. Position *
    tMmi2SpsInfo.wSytstemCheckStationModellaktiv       := HMI_GetWORD(ADR(tSpsMessage.awDaten[11])); // Hinweis: die evtl. auf der Station/Shuttle befindliche Scheibe ist ein Modell
    tMmi2SpsInfo.rSystemCheckModellVersatzVorne        := HMI_GetREAL(ADR(tSpsMessage.awDaten[12])); // Modellversatz
    tMmi2SpsInfo.rSystemCheckModellVersatzHinten       := HMI_GetREAL(ADR(tSpsMessage.awDaten[14])); // Modellversatz
    tMmi2SpsInfo.wSystemCheckScheibenDicke             := HMI_GetWORD(ADR(tSpsMessage.awDaten[16])); // Glasdicke ist binär, da für mehrere Wände die Dicke mit gegeben werden muss. Glas bis 13mm = 0 / Glasdicke > 13mm = 1
    tMmi2SpsInfo.rSystemcheckGlasGewicht               := HMI_GetREAL(ADR(tSpsMessage.awDaten[18])); // Glasgewicht, errechnet vom MMI

    // Die Wandnummer wird Bitcodiert übergeben. In der SPS wird sie aber Dezimal benötigt
    // Wand 3
    IF tMmi2SpsInfo.wSystemCheckStationSlot = 4 THEN
      tMmi2SpsInfo.wSystemCheckStationSlot := 3;
    END_IF
    // Wand 4
    IF tMmi2SpsInfo.wSystemCheckStationSlot = 8 THEN
      tMmi2SpsInfo.wSystemCheckStationSlot := 4;
    END_IF

  // MSG 69
  // Anfrage der Oberflaeche um die aktuelle Shuttleposition zu bekommen
  SB0_MMI_GETSORTIERUNGSHUTTLEPOS:
    M_SB0_MMI_GETSORTIERUNGSHUTTLEPOS := TRUE;

  // MSG 70
  // Anzeige der IO´s im MMI Service  WORT 0: 1 = sichtbar / 0 = unsichtbar
  SB0_MMI_IOANZEIGE_AKTIVIEREN_DEAKTIVIEREN:
    M_SB0_MMI_IOANZEIGE_AKTIVIEREN_DEAKTIVIEREN := TRUE;
    tMmi2SpsInfo.wlIOsAnzeigeAktivierenDeaktivieren := HMI_GetWORD(ADR(tSpsMessage.awDaten[0]));

  // MSG 71
  // Uebergabe der Auftragsdaten von der HMI fuer die Fremdanlage
  SB0_MMI_AUFTRAGSDATEN_FREMDANLAGE:
    tMmi2SpsInfo.wFremdanlageNr       := HMI_GetWORD(ADR(tSpsMessage.awDaten[0]));
    tMmi2SpsInfo.wNachrichtenIndex    := HMI_GetWORD(ADR(tSpsMessage.awDaten[1]));
    tMmi2SpsInfo.wNachrichtenAnzahl   := HMI_GetWORD(ADR(tSpsMessage.awDaten[2]));
    tMmi2SpsInfo.wScheibenanzahl      := HMI_GetWORD(ADR(tSpsMessage.awDaten[3]));
    tMmi2SpsInfo.adwScheibenID_1[0]   := HMI_GetDWORD(ADR(tSpsMessage.awDaten[4]));
    tMmi2SpsInfo.adwScheibenID_1[1]   := HMI_GetDWORD(ADR(tSpsMessage.awDaten[6]));
    tMmi2SpsInfo.adwScheibenID_1[2]   := HMI_GetDWORD(ADR(tSpsMessage.awDaten[8]));
    tMmi2SpsInfo.adwScheibenID_1[3]   := HMI_GetDWORD(ADR(tSpsMessage.awDaten[10]));
    tMmi2SpsInfo.adwScheibenID_2[0]   := HMI_GetDWORD(ADR(tSpsMessage.awDaten[12]));
    tMmi2SpsInfo.adwScheibenID_2[1]   := HMI_GetDWORD(ADR(tSpsMessage.awDaten[14]));
    tMmi2SpsInfo.adwScheibenID_2[2]   := HMI_GetDWORD(ADR(tSpsMessage.awDaten[16]));
    tMmi2SpsInfo.adwScheibenID_2[3]   := HMI_GetDWORD(ADR(tSpsMessage.awDaten[18]));
    tMmi2SpsInfo.adwScheibenID_3[0]   := HMI_GetDWORD(ADR(tSpsMessage.awDaten[20]));
    tMmi2SpsInfo.adwScheibenID_3[1]   := HMI_GetDWORD(ADR(tSpsMessage.awDaten[22]));
    tMmi2SpsInfo.adwScheibenID_3[2]   := HMI_GetDWORD(ADR(tSpsMessage.awDaten[24]));
    tMmi2SpsInfo.adwScheibenID_3[3]   := HMI_GetDWORD(ADR(tSpsMessage.awDaten[26]));

    M_SB0_MMI_AUFTRAGSDATEN_FREMDANLAGE := TRUE;

  // MSG 72
  // Auftragsinformationen waehrend der Querfahrt uebertragen
  SB0_MMI_SHUTTLE_INFORMATION:
    tMmi2SpsInfo.wAuftrag_ShuttleNummer   := HMI_GetWORD(ADR(tSpsMessage.awDaten[0]));
    tMmi2SpsInfo.rAuftrag_Laenge          := HMI_GetReal(ADR(tSpsMessage.awDaten[1]));
    tMmi2SpsInfo.wAuftrag_TranferStation  := HMI_GetWORD(ADR(tSpsMessage.awDaten[3]));
    tMmi2SpsInfo.wAuftrag_Modus           := HMI_GetWORD(ADR(tSpsMessage.awDaten[4]));
    tMmi2SpsInfo.wAuftrag_ShuttleWand     := HMI_GetWORD(ADR(tSpsMessage.awDaten[5]));
    tMmi2SpsInfo.rAuftrag_Dicke           := WORD_TO_REAL(HMI_GetWORD(ADR(tSpsMessage.awDaten[6])));
    tMmi2SpsInfo.wAuftrag_TransferWand    := HMI_GetWORD(ADR(tSpsMessage.awDaten[7]));
    // tMmi2SpsInfo.rAuftrag_Dicke           := HMI_GetReal(ADR(tSpsMessage.awDaten[8]));

    M_SB0_MMI_SHUTTLE_INFORMATION := TRUE;

  // MSG 76
  (* Hinweis:
     - Speicherfachvalidierung mittels Transfershuttle wenn ein Sensor von diesem nicht frei gefahren werden konnte
       bzw. der Einlauf- oder Aulauf- Sensor belegt wurde. Aktin ist dem SystemCheck vorgelagert (Anlage muss ich im Hand-Modus
       befinden
  *)
  SB0_MMI_TRANSFERSHUTTLECHECK:

    tMmi2SpsInfo.wTransfershuttle_Nummer1       := HMI_GetWORD(ADR(tSpsMessage.awDaten[0])); // HINWEIS: Transfer - Shuttlenummer
    tMmi2SpsInfo.wTransfershuttle_Nummer2       := HMI_GetWORD(ADR(tSpsMessage.awDaten[1])); // HINWEIS: Transfer - Shuttlenummer
    tMmi2SpsInfo.wTransfershuttle_GlasDicke     := HMI_GetWORD(ADR(tSpsMessage.awDaten[2])); // HINWEIS: Unterteilung welche Luftabfrage genommen werden muss
    tMmi2SpsInfo.rTransfershuttle_SollPosition1 := HMI_GetReal(ADR(tSpsMessage.awDaten[3])); // HINWEIS: Soll-Position des Transfershuttles
    tMmi2SpsInfo.rTransfershuttle_SollPosition2 := HMI_GetReal(ADR(tSpsMessage.awDaten[5])); // HINWEIS: Soll-Position des Transfershuttles

    M_SB0_MMI_TRANSFERSHUTTLECHECK := TRUE;

    // MSG 77/100
    // Testen der Transfershuttlepositionen
    SB0_MMI_TRANSFERSHUTTLEBUFFERSLOTCHECK,
      SB0_MMI_LIFTTRANSFERSHUTTLE:
    IF ( NOT FachkontrolleTransfershuttle.bpStarteFachkontrolle ) THEN
      FachkontrolleTransfershuttle.bpStarteFachkontrolle := TRUE;
      FachkontrolleTransfershuttle.wpStationNumber       := HMI_GetWORD(ADR(tSpsMessage.awDaten[0]));;
      FachkontrolleTransferShuttle.wpSpeicherNr          := HMI_GetWORD(ADR(tSpsMessage.awDaten[1]));
      FachkontrolleTransferShuttle.wpFachNr              := HMI_GetWORD(ADR(tSpsMessage.awDaten[2]));
      FachkontrolleTransfershuttle.rpPosition            := HMI_GetReal(ADR(tSpsMessage.awDaten[3]));
    END_IF

  // MSG 81
  SB0_MMI_RESET_ETHERCAT:
    M_SB0_MMI_RESET_ETHERCAT := TRUE;

  // MSG 99
  SB0_MMI_WATCHDOGTEST:
    tMmi2SpsInfo.wWatchDogTestCount  := HMI_GetWORD(ADR(tSpsMessage.awDaten[0]));
    M_SB0_MMI_WATCHDOGTEST := TRUE;

  // MSG 101
  // Neue Nachricht für Aufträge aller Stationen und Shuttle
  SB0_MMI_SHEET_ORDER:
    tMmi2SpsInfo.wStationsNr                             := HMI_GetWORD(ADR(tSpsMessage.awDaten[0]));         // Stationsnummer der Quellstation
    tMmi2SpsInfo.rStationsPosition                       := HMI_GetREAL(ADR(tSpsMessage.awDaten[1]));  // Stationsposition der Quellstation
    tMmi2SpsInfo.rAuftragsLaenge                         := HMI_GetREAL(ADR(tSpsMessage.awDaten[3]));  // Länge der Scheibe/Batch
    tMmi2SpsInfo.rAuftragsHoehe                          := HMI_GetREAL(ADR(tSpsMessage.awDaten[5]));  // Höhe der Scheibe/Batch
    tMmi2SpsInfo.rAuftragsDicke                          := HMI_GetREAL(ADR(tSpsMessage.awDaten[7]));  // Dicke der Scheibe/Batch
    tMmi2SpsInfo.rModellVersatzVorne                     := HMI_GetREAL(ADR(tSpsMessage.awDaten[9]));
    tMmi2SpsInfo.rModellversatzHinten                    := HMI_GetREAL(ADR(tSpsMessage.awDaten[11]));
    tMmi2SpsInfo.wErsteLetzteScheibe                     := HMI_GetWORD(ADR(tSpsMessage.awDaten[13]));         // Kennzeichnung Erste und Letzte Scheibe
    tMmi2SpsInfo.wAuftragsWand                           := HMI_GetWORD(ADR(tSpsMessage.awDaten[14]));         // Stationswand der Quellstation
    tMmi2SpsInfo.wAnzahlScheiben                         := HMI_GetWORD(ADR(tSpsMessage.awDaten[15]));         // Anzahl der Scheiben
    tMmi2SpsInfo.wAuftragsTyp                            := HMI_GetWORD(ADR(tSpsMessage.awDaten[16]));         // Auftragstyp Eintransport, Austransport, etc.
    tMmi2SpsInfo.wTransferstationsNr1                    := HMI_GetWORD(ADR(tSpsMessage.awDaten[17]));         // Stationsnummer der Zielstation 1
    tMmi2SpsInfo.wTransferstationsNr2                    := HMI_GetWORD(ADR(tSpsMessage.awDaten[18]));         // Stationsnummer der Zielstation 2
    tMmi2SpsInfo.rTransferposition1                      := HMI_GetREAL(ADR(tSpsMessage.awDaten[19]));  // Stationsposition der Zielstation 1
    tMmi2SpsInfo.rTransferposition2                      := HMI_GetREAL(ADR(tSpsMessage.awDaten[21]));  // Stationsposition der Zielstation 2
    tMmi2SpsInfo.wTransferwand                           := HMI_GetWORD(ADR(tSpsMessage.awDaten[23]));         // Stationswand der Zielstationen (1Byte = Station 1, 2Byte = Station 2)

    tMmi2SpsInfo.wNachrichtenAnzahl := HMI_GetWORD(ADR(tSpsMessage.awDaten[15]));
    tMmi2SpsInfo.wNachrichtenIndex  := HMI_GetWORD(ADR(tSpsMessage.awDaten[28]));

    IF    ( tMmi2SpsInfo.wStationsNr >= cERSTE_STATION )
    THEN
      M_SB0_MMI_SHEET_ORDER_STATION := TRUE;
    ELSE
      M_SB0_MMI_SHEET_ORDER_SHUTTLE := TRUE;
    END_IF

  // MSG 102
  // Override fuer alle Antriebe [0..100 %], Auswertung in Antriebe.prg
  SB0_MMI_DRIVEOVERRIDE:
    tMmi2SpsInfo.wMmi2SpsOverrideValue := HMI_GetWORD(ADR(tSpsMessage.awDaten[0]));
    M_SB0_MMI_DRIVEOVERRIDE := TRUE;

  // MSG 110
  // Funktion zum zurueckfahren der Glaeser und neu Positionieren im Speicher
  SB0_MMI_TS_REPOSITIONING_LITES:
    tMmi2SpsInfo.wStationsNr          := HMI_GetWORD(ADR(tSpsMessage.awDaten[0]));  // Stationsnummer der Quellstation
    tMmi2SpsInfo.rStationsPosition    := HMI_GetREAL(ADR(tSpsMessage.awDaten[1]));  // Stationsposition der Quellstation
    tMmi2SpsInfo.wTransferstationsNr1 := HMI_GetWORD(ADR(tSpsMessage.awDaten[3]));
    tMmi2SpsInfo.rTransferposition1   := HMI_GetREAL(ADR(tSpsMessage.awDaten[4]));  // Stationsposition der Quellstation
    tMmi2SpsInfo.rModellversatzHinten := HMI_GetREAL(ADR(tSpsMessage.awDaten[6]));
    tMmi2SpsInfo.rAuftragsDicke       := HMI_GetREAL(ADR(tSpsMessage.awDaten[8]));  // Dicke der Scheibe/Batch

    M_SB0_MMI_TS_REPOSITIONING_LITES := TRUE;

  ELSE

    MsgInterpret := FALSE;
    RETURN;

END_CASE

MsgInterpret := TRUE;
END_FUNCTION

(* ---- MsgToMmi.fn.st ---- *)
(* METADATA
{
	"v3Meta": {
		"objectGuid": "db865b54-9f7d-484b-b18c-e3bd89594534"
	}
}
*)
FUNCTION MsgToMmi : BOOL
// ------ Senden von Nachrichten zum MMI ------
VAR_INPUT
  auftragsnr_w: WORD;
END_VAR
VAR
  msg_st  : SpsMessage;

  wlIndex : WORD;

  wlAnzahl, wlWert, wlBenoetigt : WORD;
END_VAR
CASE( auftragsnr_w ) OF

    // Aktive Handfunktionen: Stationsnummer, niedriges Word, hohes Word.
    SB0_SPS_HANDFUNKTION_STATUS,
      SB0_SPS_SHUTTLEHANDFUNKTION_STATUS:
    msg_st.wAuftrag := auftragsnr_w;
    msg_st.wLaenge := 6;
    HMI_PutWORD(  pbyAddr := ADR( msg_st.awDaten[0] ), wVal := wSps2MmiStationsNummer );
    HMI_PutDWORD( pbyAddr := ADR( msg_st.awDaten[1] ), dwVal := dwSps2MmiHandfunktionenStatus );

  (* Hinweis:
     - Versionsstring
  *)
  SB0_SPS_SPSVERSION:
    msg_st.wAuftrag := auftragsnr_w;
    msg_st.wLaenge := INT_TO_WORD(LEN(sSpsVersion) + 1);
  // HMI_PutString( pbyAddr := ADR(msg_st.awDaten[0]), wVal := sSpsVersion);

  (* Hinweis:
     - Maschinen Statusmeldung
  *)
  SB0_SPS_SETBETRIEBSART:
    msg_st.wAuftrag := auftragsnr_w;
    msg_st.wLaenge := 20;
    HMI_PutWORD( pbyAddr := ADR( msg_st.awDaten[0] ), wVal := awSPS2MMIMaschineStatusWord[1] );
    HMI_PutWORD( pbyAddr := ADR( msg_st.awDaten[1] ), wVal := awSPS2MMIMaschineStatusWord[2] );
    HMI_PutWORD( pbyAddr := ADR( msg_st.awDaten[2] ), wVal := awSPS2MMIMaschineStatusWord[3] );
    HMI_PutWORD( pbyAddr := ADR( msg_st.awDaten[3] ), wVal := awSPS2MMIMaschineStatusWord[4] );
    HMI_PutWORD( pbyAddr := ADR( msg_st.awDaten[4] ), wVal := awSPS2MMIMaschineStatusWord[5] );
    HMI_PutWORD( pbyAddr := ADR( msg_st.awDaten[5] ), wVal := awSPS2MMIMaschineStatusWord[6] );
    HMI_PutWORD( pbyAddr := ADR( msg_st.awDaten[6] ), wVal := awSPS2MMIMaschineStatusWord[7] );
    HMI_PutWORD( pbyAddr := ADR( msg_st.awDaten[7] ), wVal := awSPS2MMIMaschineStatusWord[8] );
    HMI_PutWORD( pbyAddr := ADR( msg_st.awDaten[8] ), wVal := awSPS2MMIMaschineStatusWord[9] );
    HMI_PutWORD( pbyAddr := ADR( msg_st.awDaten[9] ), wVal := awSPS2MMIMaschineStatusWord[10] );
    HMI_PutWORD( pbyAddr := ADR( msg_st.awDaten[10] ), wVal := awSPS2MMIMaschineStatusWord[11] );

  (* Hinweis:
     - Quittung des Anlegeauftrages
       => Scheibe wurde vermessen und kann ins System eingebucht werden
       WORD [1] und [2] sind reserviert für Höhe
       WORD [3] und [4] sind reserviert für Länge
  *)
  SB0_SPS_SortierungQuittInputInQueue:  // Auftrag für den Anlegetisch
    msg_st.wAuftrag := auftragsnr_w;
    msg_st.wLaenge := 14;
    HMI_PutWORD( pbyAddr := ADR( msg_st.awDaten[0] ), wVal := wSps2MmiInputtableNummer );// Tischnummer
    HMI_PutDWORD( pbyAddr := ADR( msg_st.awDaten[6] ), dwVal := dwSps2MmiWartezeit );

  (* Hinweis:
     - -Event-State einer Station
  *)
  SBO_SPS_STATIONSEVENT:
    msg_st.wAuftrag := auftragsnr_w;
    msg_st.wLaenge := 2;
    HMI_PutWORD( pbyAddr := ADR( msg_st.awDaten[0] ), wVal := wSps2MmiStationsNummer );// Stationsnummer
    HMI_PutWORD( pbyAddr := ADR( msg_st.awDaten[1] ), wVal := wSPS2MMIStationEventStatus );// Station Event-Typ

  SB0_SPS_ErrorMSG:
    msg_st.wAuftrag := auftragsnr_w;  // Konstanten Nr. !!
    msg_st.wLaenge := 10;
    HMI_PutWORD( pbyAddr := ADR( msg_st.awDaten[0] ), wVal := wSps2MmiErrorNumber );// + Parameter z.B.: Fehlernummer des Antriebes
    HMI_PutWORD( pbyAddr := ADR( msg_st.awDaten[1] ), wVal := wSps2MmiErrorShuttleNumber );// + Parameter z.B.: Shuttlenummer
    HMI_PutWORD( pbyAddr := ADR( msg_st.awDaten[2] ), wVal := wSps2MmiErrorShuttleSchritt );// + Parameter z.B.: Schrittkettenschritt
    HMI_PutWORD( pbyAddr := ADR( msg_st.awDaten[3] ), wVal := wSps2MmiErrorShuttlePosition4 );
    HMI_PutWORD( pbyAddr := ADR( msg_st.awDaten[4] ), wVal := wSps2MmiErrorShuttlePosition5 );
    HMI_PutWORD( pbyAddr := ADR( msg_st.awDaten[5] ), wVal := wSps2MmiErrorShuttlePosition6 );
    HMI_PutWORD( pbyAddr := ADR( msg_st.awDaten[6] ), wVal := wSps2MmiErrorShuttlePosition7 );
    HMI_PutWORD( pbyAddr := ADR( msg_st.awDaten[7] ), wVal := wSps2MmiErrorShuttlePosition8 );
    HMI_PutWORD( pbyAddr := ADR( msg_st.awDaten[8] ), wVal := wSps2MmiErrorShuttlePosition9 );

  SB0_SPS_DEBUG_TRACE:
    msg_st.wAuftrag := auftragsnr_w;  // Konstanten Nr. !!
    msg_st.wLaenge := 9;
    HMI_PutWORD( pbyAddr := ADR( msg_st.awDaten[0] ), wVal := wSps2MmiDebugLogWord1); // + Parameter z.B.: Fehlernummer des Antriebes
    HMI_PutWORD( pbyAddr := ADR( msg_st.awDaten[1] ), wVal := wSps2MmiDebugLogWord2); // + Parameter z.B.: Shuttlenummer
    HMI_PutWORD( pbyAddr := ADR( msg_st.awDaten[2] ), wVal := wSps2MmiDebugLogWord3); // + Parameter z.B.: Schrittkettenschritt
    HMI_PutWORD( pbyAddr := ADR( msg_st.awDaten[3] ), wVal := wSps2MmiDebugLogWord4);
    HMI_PutWORD( pbyAddr := ADR( msg_st.awDaten[4] ), wVal := wSps2MmiDebugLogWord5);
    HMI_PutWORD( pbyAddr := ADR( msg_st.awDaten[5] ), wVal := wSps2MmiDebugLogWord6);
    HMI_PutWORD( pbyAddr := ADR( msg_st.awDaten[6] ), wVal := wSps2MmiDebugLogWord7);
    HMI_PutWORD( pbyAddr := ADR( msg_st.awDaten[7] ), wVal := wSps2MmiDebugLogWord8);
    HMI_PutWORD( pbyAddr := ADR( msg_st.awDaten[8] ), wVal := wSps2MmiDebugLogWord9);

  (* Hinweis:
     - Nachricht fuer die Scheibenmessung der Stationen
  *)
  SB0_SPS_SETSHEETSONSTATION:
    // Die Wandnummer wird Bitcodiert übergeben. In der SPS wird sie aber Dezimal benötigt
    // Wand 3
    IF ( wSps2MmiMessungSlotNummer = 3) THEN
      wSps2MmiMessungSlotNummer  := 4;
    END_IF
    msg_st.wAuftrag := auftragsnr_w;
    msg_st.wLaenge := 3;
    HMI_PutWORD( pbyAddr := ADR( msg_st.awDaten[0] ), wVal := wSps2MmiMessungStationNummer );
    HMI_PutWORD( pbyAddr := ADR( msg_st.awDaten[1] ), wVal := wSps2MmiMessungSlotNummer );
    HMI_PutWORD( pbyAddr := ADR( msg_st.awDaten[2] ), wVal := INT_TO_WORD(iSps2MmiMessungScheibenanzahl) );
    HMI_PutREAL( pbyAddr := ADR( msg_st.awDaten[3] ), rVal := rSps2MmiMessungScheibenlaenge );

  (* Hinweis:
     - Auftragsquittierung fuer die Scheibenvorpositionierung im Speicher mit dem Transfershuttle
  *)
  SB0_SPS_SortierungQuittExtractionShuttleData: //
    msg_st.wAuftrag := auftragsnr_w;
    msg_st.wLaenge := 6;
    HMI_PutWORD( pbyAddr := ADR( msg_st.awDaten[0] ), wVal := wSps2MmiQuittierungVortransportStationsNr1 );
    HMI_PutWORD( pbyAddr := ADR( msg_st.awDaten[1] ), wVal := wSps2MmiQuittierungVortransportStatus );
    HMI_PutREAL( pbyAddr := ADR( msg_st.awDaten[2] ), rVal := rgSPS2MMIExtractionShuttleGefahrenerWeg );
    HMI_PutWORD( pbyAddr := ADR( msg_st.awDaten[4] ), wVal := wSps2MmiQuittierungVortransportStationsNr2 );

  SB0_SPS_SORTIERUNGQUITTUNGVONISOLINIE:
    msg_st.wAuftrag := auftragsnr_w;
    msg_st.wLaenge := 2;
    HMI_PutWORD( pbyAddr := ADR( msg_st.awDaten[0] ), wVal := wSps2MmiQuittISOLineNr );
    HMI_PutDWORD( pbyAddr := ADR( msg_st.awDaten[1] ), dwVal := dwSps2MmiWartezeit );

  (* Hinweis:
     - Transporstatus der Eckuebergabe/Anlegetisch [Scanner] zum MMI
  *)
  SB0_SPS_TRANSPORTSTATE:
    msg_st.wAuftrag := auftragsnr_w;
    msg_st.wLaenge := 7;
    HMI_PutWORD( pbyAddr := ADR( msg_st.awDaten[0] ), wVal := wSPS2MMITRANSPORTSTATE );
    HMI_PutWORD( pbyAddr := ADR( msg_st.awDaten[1] ), wVal := wSPS2MMITransportstateStation );
    HMI_PutREAL( pbyAddr := ADR( msg_st.awDaten[2] ), rVal := rSPS2MMITransportStateLenght );
    HMI_PutREAL( pbyAddr := ADR( msg_st.awDaten[4] ), rVal := rSPS2MMITransportStateHigh );
    HMI_PutWORD( pbyAddr := ADR( msg_st.awDaten[6] ), wVal := wSPS2MMITransportstateGap );

  SB0_SPS_SHEETONINPUTTABLE:
    msg_st.wAuftrag := auftragsnr_w;
    msg_st.wLaenge := 4;
    HMI_PutWORD(  pbyAddr := ADR( msg_st.awDaten[0] ), wVal  := wSps2MmiInputtableNummer );
    HMI_PutDWORD( pbyAddr := ADR( msg_st.awDaten[1] ), dwVal := dwSps2MmiWartezeit );

  SB0_SPS_TURNSTATIONPOSITION:
    msg_st.wAuftrag := auftragsnr_w;
    msg_st.wLaenge := 6;
    HMI_PutWORD(  pbyAddr := ADR( msg_st.awDaten[0] ), wVal  := wgSps2MmiDrehStation );
    HMI_PutWORD(  pbyAddr := ADR( msg_st.awDaten[1] ), wVal  := wgSps2MmiPosDrehStation );
    HMI_PutWORD(  pbyAddr := ADR( msg_st.awDaten[2] ), wVal  := wgSps2MmiOldPosDrehStation );

  SB0_SPS_SYSTEMCHECKFINISHED:
    msg_st.wAuftrag := auftragsnr_w;
    msg_st.wLaenge := 1;
    HMI_PutWORD(  pbyAddr := ADR( msg_st.awDaten[0] ), wVal  := wSps2MmiCheckArea );
    HMI_PutWORD(  pbyAddr := ADR( msg_st.awDaten[1] ), wVal  := wSps2MmiCheckSuccessful );

  SB0_SPS_SETSHEETSONSHUTTLE:
    msg_st.wAuftrag := auftragsnr_w;
    msg_st.wLaenge := 14;
    HMI_PutWORD(  pbyAddr := ADR( msg_st.awDaten[0] ), wVal  := wSps2MmiMeasureShuttleNummer );
    HMI_PutWORD(  pbyAddr := ADR( msg_st.awDaten[1] ), wVal  := wSps2MmiMessungSlotNummer );
    HMI_PutWORD(  pbyAddr := ADR( msg_st.awDaten[2] ), wVal  := INT_TO_WORD(iSps2MmiMessungScheibenanzahl) );
    FOR wlIndex:=0 TO cMaxScheibenBeiScheibenMessung DO
      HMI_PutREAL(  pbyAddr := ADR( msg_st.awDaten[(2*(wlIndex)) + 3] ), rVal  := rSps2MmiMeasureResult[wlIndex] );
    END_FOR

    // Werte zuruecksetzen
    wSps2MmiMeasureShuttleNummer  := 0;
    wSps2MmiMessungSlotNummer     := 0;
    iSps2MmiMessungScheibenanzahl := 0;

  (* Hinweis:
     - GETTER: Anfrage des Stations- Status [z.B. Status Ein-/Aus- Transport]
  *)
  SB0_SPS_GETSTATIONSTATUS:
    msg_st.wAuftrag := auftragsnr_w;
    msg_st.wLaenge := 2;
    HMI_PutWORD(  pbyAddr := ADR( msg_st.awDaten[0] ), wVal  := wSps2MmiStationsNummer );

  SB0_SPS_SHUTTLEVORABPOSITIONIERUNGUPDATE:
    msg_st.wAuftrag := auftragsnr_w;
    msg_st.wLaenge := 4;
    HMI_PutWORD( pbyAddr := ADR( msg_st.awDaten[0] ), wVal  := wSps2MmiQuittVorabShuttleNr );
    HMI_PutREAL( pbyAddr := ADR( msg_st.awDaten[1] ), rVal := rgSPS2MMIExtractionShuttlePosition );

  SB0_SPS_QUITTSHUTTLEVORABPOSITIONIERUNG:
    msg_st.wAuftrag := auftragsnr_w;
    msg_st.wLaenge := 4;
    HMI_PutWORD( pbyAddr := ADR( msg_st.awDaten[0] ), wVal := wSps2MmiQuittVorabShuttleNr );
    HMI_PutREAL( pbyAddr := ADR( msg_st.awDaten[1] ), rVal := rgSPS2MMIExtractionShuttlePosition );

  SB0_SPS_SORTIERUNGSHUTTLEPOS:
    msg_st.wAuftrag := auftragsnr_w;
    msg_st.wLaenge := 30;
    HMI_PutREAL( pbyAddr := ADR( msg_st.awDaten[0] ),  rVal := rSps2MmiShuttlePosition[0] );
    HMI_PutREAL( pbyAddr := ADR( msg_st.awDaten[2] ),  rVal := rSps2MmiShuttlePosition[1] );
    HMI_PutREAL( pbyAddr := ADR( msg_st.awDaten[4] ),  rVal := rSps2MmiShuttlePosition[2] );
    HMI_PutREAL( pbyAddr := ADR( msg_st.awDaten[6] ),  rVal := rSps2MmiShuttlePosition[3] );
    HMI_PutREAL( pbyAddr := ADR( msg_st.awDaten[8] ),  rVal := rSps2MmiShuttlePosition[4] );
    HMI_PutREAL( pbyAddr := ADR( msg_st.awDaten[10] ), rVal := rSps2MmiShuttlePosition[5] );
    HMI_PutREAL( pbyAddr := ADR( msg_st.awDaten[12] ), rVal := rSps2MmiShuttlePosition[6] );
    HMI_PutREAL( pbyAddr := ADR( msg_st.awDaten[14] ), rVal := rSps2MmiShuttlePosition[7] );
    HMI_PutREAL( pbyAddr := ADR( msg_st.awDaten[16] ), rVal := rSps2MmiShuttlePosition[8] );
    HMI_PutREAL( pbyAddr := ADR( msg_st.awDaten[18] ), rVal := rSps2MmiShuttlePosition[9] );
    HMI_PutREAL( pbyAddr := ADR( msg_st.awDaten[20] ), rVal := rSps2MmiShuttlePosition[10] );
    HMI_PutREAL( pbyAddr := ADR( msg_st.awDaten[22] ), rVal := rSps2MmiShuttlePosition[11] );

  SB0_SPS_SHUTTLEVORABPOSITIONIERUNGABBRUCH:
    msg_st.wAuftrag := auftragsnr_w;
    msg_st.wLaenge := 4;
    HMI_PutWORD(  pbyAddr := ADR( msg_st.awDaten[0] ), wVal  := wgSps2MmiShuttleNr );
    HMI_PutREAL( pbyAddr := ADR( msg_st.awDaten[1] ),  rVal := rSps2MmiPosition );
    HMI_PutWORD(  pbyAddr := ADR( msg_st.awDaten[3] ), wVal  := wSps2ShuttleStopped[wgSps2MmiShuttleNr] );

    SB0_SPS_TRANSFERSHUTTLEBUFFERSLOTPOS,
      SB0_SPS_LIFTEDTRANSFERSHUTTLEPOSITION:
    msg_st.wAuftrag := auftragsnr_w;
    msg_st.wLaenge := 6;
    HMI_PutWORD(  pbyAddr := ADR( msg_st.awDaten[0] ), wVal  := wgSps2MmiShuttleNr );
    HMI_PutREAL(  pbyAddr := ADR( msg_st.awDaten[1] ), rVal  := wSps2MmiValidierungsPosition );
    HMI_PutWORD(  pbyAddr := ADR( msg_st.awDaten[3] ), wVal  := wSps2MmiValidierungsSpeicher );
    HMI_PutWORD(  pbyAddr := ADR( msg_st.awDaten[4] ), wVal  := wSps2MmiValidierungsFach );

  SB0_SPS_SHUTTLEVORABPOSITIONIERUNGREADY:
    msg_st.wAuftrag := auftragsnr_w;
    msg_st.wLaenge := 3;
    HMI_PutWORD(  pbyAddr := ADR( msg_st.awDaten[0] ), wVal  := wSps2MmiStationsNummer );
    HMI_PutREAL(  pbyAddr := ADR( msg_st.awDaten[1] ), rVal  := rSps2MmiPosition );

  SB0_SPS_TRANSFERSHUTTLEFEHLER:
    msg_st.wAuftrag := auftragsnr_w;
    msg_st.wLaenge := 6;
    HMI_PutWORD(  pbyAddr := ADR( msg_st.awDaten[0] ), wVal  := wgSps2MmiShuttleNr );
    HMI_PutREAL(  pbyAddr := ADR( msg_st.awDaten[1] ), rVal  := rgSPS2MMIExtractionShuttlePosition );
    HMI_PutWORD(  pbyAddr := ADR( msg_st.awDaten[3] ), wVal  := wSps2MmiFehlertyp );

  SB0_SPS_TRANSFERSHUTTLECHECK_ABGESCHLOSSEN:
    msg_st.wAuftrag := auftragsnr_w;
    msg_st.wLaenge := 6;
    HMI_PutWORD(  pbyAddr := ADR( msg_st.awDaten[0] ), wVal  := wgSps2MmiShuttleNr );
    HMI_PutWORD(  pbyAddr := ADR( msg_st.awDaten[1] ), wVal  := wSps2MmiValidierungsStatus );

  SB0_SPS_FACHAUFNAHMEDATEN:
    msg_st.wAuftrag := auftragsnr_w;
    msg_st.wLaenge := 4;
    HMI_PutREAL(  pbyAddr := ADR( msg_st.awDaten[1] ), rVal  := rSPS2MMIFachaufnahmePosition );
    HMI_PutWORD(  pbyAddr := ADR( msg_st.awDaten[3] ), wVal  := wSPS2MMIFachaufnahmeAnalogwert );

  (* Hinweis:
     - Neue Nachricht zum quittieren von Aufträgen
  *)
  SB0_SPS_QUIT_SHEET_ORDER:
    msg_st.wAuftrag   := auftragsnr_w;
    msg_st.wLaenge    := 4;
    HMI_PutWORD(  pbyAddr := ADR( msg_st.awDaten[0] ),  wVal  := wSps2MmiZielStation );
    HMI_PutWORD(  pbyAddr := ADR( msg_st.awDaten[1] ),  wVal  := wSps2MmiQuellStation );
    HMI_PutWORD(  pbyAddr := ADR( msg_st.awDaten[2] ),  wVal  := wSps2MmiZielWand );
    HMI_PutWORD(  pbyAddr := ADR( msg_st.awDaten[3] ),  wVal  := wSps2MmiQuellWand );
    HMI_PutDWORD( pbyAddr := ADR( msg_st.awDaten[4] ), dwVal  := dwSps2MmiWartezeit );
    HMI_PutWORD(  pbyAddr := ADR( msg_st.awDaten[6] ),  wVal  := wSPS2MMIAuftragstyp );

  SB0_SPS_SCHNITTSTELLENDATENFREMDANLAGE:
    msg_st.wAuftrag    := auftragsnr_w;
    msg_st.wLaenge     := 4;
    HMI_PutWORD(  pbyAddr := ADR( msg_st.awDaten[0] ),  wVal  := wSps2Mmi_SationsNummer );
    HMI_PutWORD(  pbyAddr := ADR( msg_st.awDaten[1] ),  wVal  := wSps2Mmi_NachrichtenIndex );
    HMI_PutWORD(  pbyAddr := ADR( msg_st.awDaten[2] ),  wVal  := wSps2Mmi_NachrichtenAnzahl );
    HMI_PutWORD(  pbyAddr := ADR( msg_st.awDaten[3] ),  wVal  := wSps2Mmi_AnzahlScheiben );
    HMI_PutDWORD(  pbyAddr := ADR( msg_st.awDaten[4] ),  dwVal  := adwSps2Mmi_Daten_1[0] );
    HMI_PutDWORD(  pbyAddr := ADR( msg_st.awDaten[6] ),  dwVal  := adwSps2Mmi_Daten_1[1] );
    HMI_PutDWORD(  pbyAddr := ADR( msg_st.awDaten[8] ),  dwVal  := adwSps2Mmi_Daten_1[2] );
    HMI_PutDWORD(  pbyAddr := ADR( msg_st.awDaten[10] ),  dwVal  := adwSps2Mmi_Daten_1[3] );
    HMI_PutDWORD(  pbyAddr := ADR( msg_st.awDaten[12] ),  dwVal  := adwSps2Mmi_Daten_2[0] );
    HMI_PutDWORD(  pbyAddr := ADR( msg_st.awDaten[14] ),  dwVal  := adwSps2Mmi_Daten_2[1] );
    HMI_PutDWORD(  pbyAddr := ADR( msg_st.awDaten[16] ),  dwVal  := adwSps2Mmi_Daten_2[2] );
    HMI_PutDWORD(  pbyAddr := ADR( msg_st.awDaten[18] ),  dwVal  := adwSps2Mmi_Daten_2[3] );
    HMI_PutDWORD(  pbyAddr := ADR( msg_st.awDaten[20] ),  dwVal  := adwSps2Mmi_Daten_3[0] );
    HMI_PutDWORD(  pbyAddr := ADR( msg_st.awDaten[22] ),  dwVal  := adwSps2Mmi_Daten_3[1] );
    HMI_PutDWORD(  pbyAddr := ADR( msg_st.awDaten[24] ),  dwVal  := adwSps2Mmi_Daten_3[2] );
    HMI_PutDWORD(  pbyAddr := ADR( msg_st.awDaten[26] ),  dwVal  := adwSps2Mmi_Daten_3[3] );

  (* Hinweis:
     - Ausmessen von FW
  *)
  SB0_SPS_POSITIONMEASUREDATA:
    msg_st.wAuftrag := auftragsnr_w;
    msg_st.wLaenge := 5;
    HMI_PutWORD(  pbyAddr := ADR( msg_st.awDaten[0] ),  wVal  := wSps2MmiStationsNummer );
    HMI_PutREAL(  pbyAddr := ADR( msg_st.awDaten[1] ),  rVal  := rSps2MmiPosition );

  SB0_SPS_STATIONSTATUS:
    msg_st.wAuftrag := auftragsnr_w;
    msg_st.wLaenge := 2;
    HMI_PutWORD(  pbyAddr := ADR( msg_st.awDaten[0] ),  wVal  := wSps2MmiStationsNummer );
    HMI_PutWORD(  pbyAddr := ADR( msg_st.awDaten[1] ),  wVal  := wSPS2MMIStationsStatusWord1 );
    HMI_PutWORD(  pbyAddr := ADR( msg_st.awDaten[2] ),  wVal  := wSPS2MMIStationsStatusWord2 );

  SB0_SPS_SHEETREMOVEDAPPROVALWALL:
    msg_st.wAuftrag := auftragsnr_w;
    msg_st.wLaenge := 3;
    HMI_PutWORD(  pbyAddr := ADR( msg_st.awDaten[0] ),  wVal  := wSps2MmiStationsNummer );

  SB0_SPS_WATCHDOGTEST:
    msg_st.wAuftrag := auftragsnr_w;
    msg_st.wLaenge := 3;
    HMI_PutWORD(  pbyAddr := ADR( msg_st.awDaten[0] ),  wVal  := wSps2MmiWatchDogTestCount );

  // ++++++++++++++++++++++++ Fächerwagenstationen ++++++++++++++++++++++++++++++++++++
  (* Hinweis [FAECHERWAGEN]:
     - Faecherwagenwechsel von Station A nach B erfolgreich
  *)
  SB0_SPS_RACKONLOADINGSTATION:
    msg_st.wAuftrag := auftragsnr_w;
    msg_st.wLaenge := 3;
    HMI_PutWORD(  pbyAddr := ADR( msg_st.awDaten[0] ),  wVal  := wSps2MmiRackPositionNummer );
    HMI_PutWORD(  pbyAddr := ADR( msg_st.awDaten[1] ),  wVal  := wSps2MmiRackPosition );
    HMI_PutWORD(  pbyAddr := ADR( msg_st.awDaten[2] ),  wVal  := wSps2MmiRackNumber );

  (* Hinweis [FAECHERWAGEN]:
     - Anforderung zum einbuchen des Faecherwagens
        => Status: 1 = FW auf Station 1 / 2 = FW auf Station 2 / etc.
  *)
  SB0_SPS_RACKLOGIN:
    msg_st.wAuftrag := auftragsnr_w;
    msg_st.wLaenge := 2;
    HMI_PutWORD(  pbyAddr := ADR( msg_st.awDaten[0] ),  wVal  := wSps2FaecherwagenStationNr );

  SB0_SPS_SortierungRackinPos: // Fächerwagenwechsel von Station A nach B erfolgreich
    msg_st.wAuftrag := auftragsnr_w;
    msg_st.wLaenge := 2;
    HMI_PutWORD(  pbyAddr := ADR( msg_st.awDaten[0] ),  wVal  := wSps2FaecherwagenStart );// Wo kommt der Wagen her
    HMI_PutWORD(  pbyAddr := ADR( msg_st.awDaten[1] ),  wVal  := wSps2FaecherwagenStart );// Wo geht der Wagen hin

  (* Hinweis:
     - [FAECHERWAGENSTATION] Gibt den Status der Faecherwagenstation zurueck
       => 0 = wird nicht benutzt
       => 1 = frei
       => 2 = belegt
       Wichtig:
       => Groesse des Arrays <awSps2MmmiStatusFaecherwagenstation> beachten ggf. den Index vergroessern
       => <igIndexFaecherwagenDatenSenden> Aufgrund des Datenwortes das bei "0" startet [Index]
  *)

  (* Hinweis [FAECHERWAGEN]:
     - Anforderung zum einbuchen des Faecherwagens
        => Status: 1 = FW auf Station 1 / 2 = FW auf Station 2 / etc.
  *)
  SB0_SPS_RACKPOSITION:
    msg_st.wAuftrag := auftragsnr_w;
    msg_st.wLaenge := 4;
    HMI_PutWORD(  pbyAddr := ADR( msg_st.awDaten[0] ),  wVal  := wSps2MmiRackPositionNummer );
    HMI_PutWORD(  pbyAddr := ADR( msg_st.awDaten[1] ),  wVal  := wSps2MmiRackPosition );
    HMI_PutWORD(  pbyAddr := ADR( msg_st.awDaten[2] ),  wVal  := wSps2MmiRackNumber );

  SB0_SPS_SETSTATUSLOADINGSTATIONS:
    msg_st.wAuftrag := auftragsnr_w;
    msg_st.wLaenge := 10;

    igIndexFaecherwagenDatenSenden := 0;

    FOR wlIndex := 0 TO 29 DO
      HMI_PutWORD(  pbyAddr := ADR( msg_st.awDaten[igIndexFaecherwagenDatenSenden] ),  wVal  := awSps2MmiStatusFaecherwagenstationen[igIndexFaecherwagenDatenSenden] );
      igIndexFaecherwagenDatenSenden := igIndexFaecherwagenDatenSenden + 1;
    END_FOR

  SB0_SPS_SORTIERUNGRACKSTATIONSTATUS:
    msg_st.wAuftrag := auftragsnr_w;
    msg_st.wLaenge := 4;
    HMI_PutWORD(  pbyAddr := ADR( msg_st.awDaten[0] ),  wVal  := wSps2MmiRackNumber );
    HMI_PutWORD(  pbyAddr := ADR( msg_st.awDaten[1] ),  wVal  := wSps2MmiRackStatus );// 1 Wagen wird ausgeschleust, 2 Wagen wird Notausgeschleust

  //  - Anfrage vom MMI nach dem Status einer EINZELNEN Fächerwagenstation => belegt, Muting OK, RFID-Nr.
  SB0_SPS_STATUSRACKSTATION:
    msg_st.wAuftrag := auftragsnr_w;
    msg_st.wLaenge := 6;
    HMI_PutWORD(  pbyAddr := ADR( msg_st.awDaten[0] ),  wVal  := INT_TO_WORD(igRackStationNumber) );
    HMI_PutWORD(  pbyAddr := ADR( msg_st.awDaten[1] ),  wVal  := wgRackPresent );
    HMI_PutWORD(  pbyAddr := ADR( msg_st.awDaten[2] ),  wVal  := INT_TO_WORD(igRackNumber) );

  (* Hinweis:
     - Generisches Stations-Update: [0] Station, [1] Updatetyp, [2] Anzahl Werte, danach je Wert: Datentyp + Wert
  *)
  SB0_SPS_STATION_UPDATE:
    msg_st.wAuftrag := auftragsnr_w;
    HMI_PutWORD( pbyAddr := ADR( msg_st.awDaten[0] ), wVal := stStationUpdate.wStationsNummer );
    HMI_PutWORD( pbyAddr := ADR( msg_st.awDaten[1] ), wVal := TO_WORD( stStationUpdate.eUpdateTyp ) );
    wlIndex  := 3;
    wlAnzahl := 0;
    FOR wlWert := 1 TO MIN( stStationUpdate.wAnzahlWerte, 13 ) DO
      // Platzbedarf in Words inkl. Datentyp-Word
      CASE stStationUpdate.astWerte[wlWert].eDatenTyp OF
        UpdateDatenTyp_EN.TYP_WORD, UpdateDatenTyp_EN.TYP_BOOL: wlBenoetigt := 2;
        UpdateDatenTyp_EN.TYP_DWORD, UpdateDatenTyp_EN.TYP_REAL: wlBenoetigt := 3;
        ELSE
          wlBenoetigt := 0;
      END_CASE
      IF ( wlBenoetigt = 0 ) OR ( wlIndex + wlBenoetigt > 30 ) THEN
        EXIT;
      END_IF

      HMI_PutWORD( pbyAddr := ADR( msg_st.awDaten[wlIndex] ), wVal := TO_WORD( stStationUpdate.astWerte[wlWert].eDatenTyp ) );
      CASE stStationUpdate.astWerte[wlWert].eDatenTyp OF
        UpdateDatenTyp_EN.TYP_WORD:  HMI_PutWORD(  pbyAddr := ADR( msg_st.awDaten[wlIndex + 1] ), wVal  := stStationUpdate.astWerte[wlWert].wWert );
        UpdateDatenTyp_EN.TYP_DWORD: HMI_PutDWORD( pbyAddr := ADR( msg_st.awDaten[wlIndex + 1] ), dwVal := stStationUpdate.astWerte[wlWert].dwWert );
        UpdateDatenTyp_EN.TYP_REAL:  HMI_PutREAL(  pbyAddr := ADR( msg_st.awDaten[wlIndex + 1] ), rVal  := stStationUpdate.astWerte[wlWert].rWert );
        UpdateDatenTyp_EN.TYP_BOOL:  HMI_PutWORD(  pbyAddr := ADR( msg_st.awDaten[wlIndex + 1] ), wVal  := SEL( stStationUpdate.astWerte[wlWert].bWert, 0, 1 ) );
      END_CASE
      wlIndex  := wlIndex + wlBenoetigt;
      wlAnzahl := wlAnzahl + 1;
    END_FOR
    HMI_PutWORD( pbyAddr := ADR( msg_st.awDaten[2] ), wVal := wlAnzahl ); // tatsaechlich gesendete Werte
    msg_st.wLaenge := wlIndex * 2;                                        // Laenge in Byte

  ELSE
    MsgToMmi := FALSE;
    RETURN;
END_CASE;

TCPMain.l_fb_SortjetHMI.PutMsg( smpSpsMessage := msg_st, bpTrig := FALSE );
MsgToMmi := TRUE;
END_FUNCTION

(* ---- SocketIsReadable.fn.st ---- *)
(* METADATA
{
	"v3Meta": {
		"objectGuid": "0cffa44a-96d6-4cd8-9f3c-3120d05aae22"
	}
}
*)
FUNCTION SocketIsReadable : UDINT
//  Function to detect if data for reading is available on socket.
//  Return: Availability of data
VAR_INPUT
  hSocket: RTS_IEC_HANDLE; // Socket-ID
  diTimeout : DINT; // Timeout in ms
END_VAR
VAR
  fdRead: SysSocket.SOCKET_FD_SET;
  tvTimeout: SysSocket.SOCKET_TIMEVAL;
  diSysSockSelect_Return : UDINT;
  diReadySockets : DINT;
END_VAR

tvTimeout.tv_sec := diTimeout / 1000;
tvTimeout.tv_usec := (diTimeout MOD 1000) * 1000;
fdRead.fd_count := 1;
fdRead.fd_array[0] := hSocket;

diReadySockets := 0;
diSysSockSelect_Return := SysSockSelect(UDINT_TO_DINT(fdRead.fd_count), ADR(fdRead), 0, 0, ADR(tvTimeout), ADR(diReadySockets));
IF diSysSockSelect_Return = CmpErrors.Errors.ERR_OK THEN
  IF diReadySockets > 0 THEN
    SocketIsReadable := 1;
  ELSE
    SocketIsReadable := 0;
  END_IF
ELSE
  SocketIsReadable := 0;
END_IF
END_FUNCTION

(* ---- TcpReceiveData.fn.st ---- *)
(* METADATA
{
	"v3Meta": {
		"objectGuid": "b74d4ba4-35aa-49dc-9263-31d6cf99974e"
	}
}
*)
FUNCTION TcpReceiveData : __XINT
//  Receive data from a TCP socket.
//  Return: Number of bytes received or a value < 0 for an error (-1: gracefully closed; -2: error)
VAR_INPUT
  diSocket: RTS_IEC_HANDLE; // Socket-ID
  pbyData: POINTER TO DWORD; // Address of data buffer
  diDataSize: DINT; // Size of data to receive
  diTimeout: DINT; // Timeout in ms
  tcpLastError : POINTER TO LINT;
END_VAR
VAR
END_VAR

TcpReceiveData := 0;

IF SocketIsReadable(diSocket, diTimeout) > 0 THEN
  TcpReceiveData := SysSockRecv(diSocket, pbyData, diDataSize, 0,0); // Returns 0 if gracefully closed or -1 for an error
  IF TcpReceiveData <= 0 THEN
    TcpReceiveData := (*TcpReceiveData*) - 1;
    IF tcpLastError^ = 0 THEN
      tcpLastError^ := TcpReceiveData;
    END_IF
  END_IF
END_IF
END_FUNCTION

(* ---- TcpSendData.fn.st ---- *)
(* METADATA
{
	"v3Meta": {
		"objectGuid": "c3a65185-b6f7-4978-83ae-2e8140594d8c"
	}
}
*)
FUNCTION TcpSendData : __XINT
//  Send data via TCP socket.
//  Return: Number of bytes sent or a value < 0 for an error (-1: gracefully closed; -2: error)
VAR_INPUT
  diSocket: RTS_IEC_HANDLE; // Socket-ID
  pbyData: POINTER TO DWORD; // Address of data buffer
  diDataSize: DINT; // Size of data to send
  tcpLastError : POINTER TO LINT;
END_VAR
VAR
  iecResult : RTS_IEC_RESULT;
END_VAR

TcpSendData := SysSockSend(diSocket, pbyData, diDataSize, SOCKET_MSG_DONTWAIT, ADR(iecResult));
IF iecResult = CmpErrors.Errors.ERR_SOCK_WOULDBLOCK THEN
  TcpSendData := 0;
ELSE
  IF TcpSendData < 0 AND TcpSendData <> -6 AND TcpSendData <> -1 THEN
    TcpSendData := (*TcpSendData*) - 1;

    IF tcpLastError^ = 0 THEN
      tcpLastError^ := TcpSendData;
    END_IF
  END_IF
END_IF
END_FUNCTION

(* ---- TcpServerOpenSocket.fn.st ---- *)
(* METADATA
{
	"v3Meta": {
		"objectGuid": "36dfe783-e7c1-434c-babf-2b0976501267"
	}
}
*)
FUNCTION TcpServerOpenSocket : RTS_IEC_HANDLE
//  Opens a TCP server socket.
//  Return: Socket-ID
VAR_INPUT
  uiPort: UINT; // Port number
  diMaxConnections: DINT; // Max possible client connections of the server
END_VAR
VAR
  hSocket: RTS_IEC_HANDLE;
  pResult: RTS_IEC_RESULT;
  uiResult: UDINT;
  uiCloseResult: UDINT;
  sa: SOCKADDRESS;
  dwValue: DWORD := 1;
END_VAR

hSocket := SysSockCreate(SOCKET_AF_INET, SOCKET_STREAM, SOCKET_IPPROTO_TCP, ADR(pResult));

IF hSocket <> RTS_INVALID_HANDLE THEN
  SysSockSetOption(hSocket, SOCKET_SOL, SOCKET_SO_REUSEADDR, ADR(dwValue), SIZEOF(dwValue));
  sa.sin_family     := SOCKET_AF_INET;
  sa.sin_addr.ulAddr := SOCKET_INADDR_ANY;
  sa.sin_port       := SysSockHtons(uiPort);
  uiResult       := SysSockBind(hSocket, ADR(sa), SIZEOF(sa));

  IF uiResult <> CmpErrors.Errors.ERR_OK THEN
    uiCloseResult := SysSockClose(hSocket);
    hSocket := RTS_INVALID_HANDLE;
  ELSE
    uiResult := SysSockListen(hSocket, diMaxConnections);
    IF uiResult <> CmpErrors.Errors.ERR_OK THEN
      uiCloseResult := SysSockClose(hSocket);
      hSocket := RTS_INVALID_HANDLE;
    END_IF
  END_IF
END_IF
TcpServerOpenSocket := hSocket;
END_FUNCTION

(* ---- TcpServerWaitForConnect.fn.st ---- *)
(* METADATA
{
	"v3Meta": {
		"objectGuid": "244699a7-7b28-4ca6-ad52-b215d0417df3"
	}
}
*)
FUNCTION TcpServerWaitForConnect : TCP_CLIENT_ACCEPT
//  Wait for a client to connect.
//  Return: Socket and IP-Address of connected client
VAR_INPUT
  hSocket: RTS_IEC_HANDLE; // Socket-ID
  diTimeout: DINT; // Timeout in ms
END_VAR
VAR
  pResult: RTS_IEC_RESULT;
  sa: SOCKADDRESS;
  ia: INADDR;
  diSize: DINT;
END_VAR

TcpServerWaitForConnect.hSocket := RTS_INVALID_HANDLE;
TcpServerWaitForConnect.stIPAddress := '';

IF SocketIsReadable(hSocket, diTimeout) > 0 THEN
  diSize := SIZEOF(sa);
  TcpServerWaitForConnect.hSocket := SysSockAccept(hSocket, ADR(sa), ADR(diSize),ADR(pResult));
  IF TcpServerWaitForConnect.hSocket <> RTS_INVALID_HANDLE THEN
    ia.ulAddr := sa.sin_addr.ulAddr;
    SysSockInetNtoa(ADR(ia), TcpServerWaitForConnect.stIPAddress, SIZEOF(TcpServerWaitForConnect.stIPAddress));
  END_IF
END_IF
END_FUNCTION

(* ---- Hegla_Gateway_Komm_FB.fb.st ---- *)
(* METADATA
{
	"v3Meta": {
		"objectGuid": "1190007f-e857-4ecd-9ce5-2fcdfdbf097c"
	}
}
*)
FUNCTION_BLOCK Hegla_Gateway_Komm_FB
VAR_INPUT

  SpsToMmi    : SPSTOMMI;
  MmiToSps    : MMITOSPS;

END_VAR
VAR_OUTPUT

  o_b_ConnectionStart : BOOL;
  o_b_WatchdogOk : BOOL;

END_VAR
VAR
  tonlOpenForClient : TON;

  smqSpsMessageQueue : SpsMessageQueue;

  tcpLastError : LINT;
  tcpTrace : INT;

  bgTcpConnected : BOOL;

  // MMI->SPS
  MmiToSpsMem : MMITOSPS;

  // SPS->MMI
  SpsToMmiMem : SPSTOMMI;

  // Datentabelle für die CRC32-Prüfsummenberechnung
  adwgCrcTable : ARRAY[0..255] OF DWORD := [16#00000000, 16#77073096, 16#EE0E612C, 16#990951BA,
                                             16#076DC419, 16#706AF48F, 16#E963A535, 16#9E6495A3,
                                             16#0EDB8832, 16#79DCB8A4, 16#E0D5E91E, 16#97D2D988,
                                             16#09B64C2B, 16#7EB17CBD, 16#E7B82D07, 16#90BF1D91,
                                             16#1DB71064, 16#6AB020F2, 16#F3B97148, 16#84BE41DE,
                                             16#1ADAD47D, 16#6DDDE4EB, 16#F4D4B551, 16#83D385C7,
                                             16#136C9856, 16#646BA8C0, 16#FD62F97A, 16#8A65C9EC,
                                             16#14015C4F, 16#63066CD9, 16#FA0F3D63, 16#8D080DF5,
                                             16#3B6E20C8, 16#4C69105E, 16#D56041E4, 16#A2677172,
                                             16#3C03E4D1, 16#4B04D447, 16#D20D85FD, 16#A50AB56B,
                                             16#35B5A8FA, 16#42B2986C, 16#DBBBC9D6, 16#ACBCF940,
                                             16#32D86CE3, 16#45DF5C75, 16#DCD60DCF, 16#ABD13D59,
                                             16#26D930AC, 16#51DE003A, 16#C8D75180, 16#BFD06116,
                                             16#21B4F4B5, 16#56B3C423, 16#CFBA9599, 16#B8BDA50F,
                                             16#2802B89E, 16#5F058808, 16#C60CD9B2, 16#B10BE924,
                                             16#2F6F7C87, 16#58684C11, 16#C1611DAB, 16#B6662D3D,
                                             16#76DC4190, 16#01DB7106, 16#98D220BC, 16#EFD5102A,
                                             16#71B18589, 16#06B6B51F, 16#9FBFE4A5, 16#E8B8D433,
                                             16#7807C9A2, 16#0F00F934, 16#9609A88E, 16#E10E9818,
                                             16#7F6A0DBB, 16#086D3D2D, 16#91646C97, 16#E6635C01,
                                             16#6B6B51F4, 16#1C6C6162, 16#856530D8, 16#F262004E,
                                             16#6C0695ED, 16#1B01A57B, 16#8208F4C1, 16#F50FC457,
                                             16#65B0D9C6, 16#12B7E950, 16#8BBEB8EA, 16#FCB9887C,
                                             16#62DD1DDF, 16#15DA2D49, 16#8CD37CF3, 16#FBD44C65,
                                             16#4DB26158, 16#3AB551CE, 16#A3BC0074, 16#D4BB30E2,
                                             16#4ADFA541, 16#3DD895D7, 16#A4D1C46D, 16#D3D6F4FB,
                                             16#4369E96A, 16#346ED9FC, 16#AD678846, 16#DA60B8D0,
                                             16#44042D73, 16#33031DE5, 16#AA0A4C5F, 16#DD0D7CC9,
                                             16#5005713C, 16#270241AA, 16#BE0B1010, 16#C90C2086,
                                             16#5768B525, 16#206F85B3, 16#B966D409, 16#CE61E49F,
                                             16#5EDEF90E, 16#29D9C998, 16#B0D09822, 16#C7D7A8B4,
                                             16#59B33D17, 16#2EB40D81, 16#B7BD5C3B, 16#C0BA6CAD,
                                             16#EDB88320, 16#9ABFB3B6, 16#03B6E20C, 16#74B1D29A,
                                             16#EAD54739, 16#9DD277AF, 16#04DB2615, 16#73DC1683,
                                             16#E3630B12, 16#94643B84, 16#0D6D6A3E, 16#7A6A5AA8,
                                             16#E40ECF0B, 16#9309FF9D, 16#0A00AE27, 16#7D079EB1,
                                             16#F00F9344, 16#8708A3D2, 16#1E01F268, 16#6906C2FE,
                                             16#F762575D, 16#806567CB, 16#196C3671, 16#6E6B06E7,
                                             16#FED41B76, 16#89D32BE0, 16#10DA7A5A, 16#67DD4ACC,
                                             16#F9B9DF6F, 16#8EBEEFF9, 16#17B7BE43, 16#60B08ED5,
                                             16#D6D6A3E8, 16#A1D1937E, 16#38D8C2C4, 16#4FDFF252,
                                             16#D1BB67F1, 16#A6BC5767, 16#3FB506DD, 16#48B2364B,
                                             16#D80D2BDA, 16#AF0A1B4C, 16#36034AF6, 16#41047A60,
                                             16#DF60EFC3, 16#A867DF55, 16#316E8EEF, 16#4669BE79,
                                             16#CB61B38C, 16#BC66831A, 16#256FD2A0, 16#5268E236,
                                             16#CC0C7795, 16#BB0B4703, 16#220216B9, 16#5505262F,
                                             16#C5BA3BBE, 16#B2BD0B28, 16#2BB45A92, 16#5CB36A04,
                                             16#C2D7FFA7, 16#B5D0CF31, 16#2CD99E8B, 16#5BDEAE1D,
                                             16#9B64C2B0, 16#EC63F226, 16#756AA39C, 16#026D930A,
                                             16#9C0906A9, 16#EB0E363F, 16#72076785, 16#05005713,
                                             16#95BF4A82, 16#E2B87A14, 16#7BB12BAE, 16#0CB61B38,
                                             16#92D28E9B, 16#E5D5BE0D, 16#7CDCEFB7, 16#0BDBDF21,
                                             16#86D3D2D4, 16#F1D4E242, 16#68DDB3F8, 16#1FDA836E,
                                             16#81BE16CD, 16#F6B9265B, 16#6FB077E1, 16#18B74777,
                                             16#88085AE6, 16#FF0F6A70, 16#66063BCA, 16#11010B5C,
                                             16#8F659EFF, 16#F862AE69, 16#616BFFD3, 16#166CCF45,
                                             16#A00AE278, 16#D70DD2EE, 16#4E048354, 16#3903B3C2,
                                             16#A7672661, 16#D06016F7, 16#4969474D, 16#3E6E77DB,
                                             16#AED16A4A, 16#D9D65ADC, 16#40DF0B66, 16#37D83BF0,
                                             16#A9BCAE53, 16#DEBB9EC5, 16#47B2CF7F, 16#30B5FFE9,
                                             16#BDBDF21C, 16#CABAC28A, 16#53B39330, 16#24B4A3A6,
                                             16#BAD03605, 16#CDD70693, 16#54DE5729, 16#23D967BF,
                                             16#B3667A2E, 16#C4614AB8, 16#5D681B02, 16#2A6F2B94,
                                             16#B40BBE37, 16#C30C8EA1, 16#5A05DF1B, 16#2D02EF8D];

  //GetMessage
  i : WORD;

  ilAuftraegeAnz       : INT := 0;
  ilAuftragIndex       : INT := 0;
  dwAuftragsChecksumme : DWORD;
  asmSpsMessage        : ARRAY[0..4] OF SpsMessage;
  smlSpsMessage        : SpsMessage;
  smlErrorMsg          : SpsMessage;

  //MessageBegin
  dwlChecksumme0 : DWORD;
  dwlChecksumme1 : DWORD;

  //MsgPoll
  smlSpsMessage_POLL : SpsMessage;

  //WatchDog
  dwlCrc32Value          : DWORD;
  dwAuftragsChecksumme_WatchDog   : DWORD;
  ildiff          : INT;
  tlTimeOut       : TIME;
  tlTimeDiff      : TIME;
  wlWatchdogOk      : WORD;
  bTimeOff        : BOOL;
  wZyklenOff      : WORD;

  hSocket: RTS_IEC_HANDLE := RTS_INVALID_HANDLE;
  Client : TCP_CLIENT_ACCEPT;

  bInit: BOOL:= TRUE;

  blVerbindungReset: BOOL;
  rtlVerbindungReset: R_TRIG;
  tnlVerbindungReset: TON;
  wlVerbindungReset: WORD := 5000;

  // ReadMsg
  diReceived   : LINT;
  bBuffer_Read : ARRAY[0..1023] OF BYTE;
  diLenght     : DINT;
  pbCunrrent   : POINTER TO BYTE;
  mhHeader     : MsgHeader;
  diRemaining  : DINT;
  j            : WORD;
  pbCurPos_Read     : POINTER TO BYTE;

  // SendMsg
  diSent        : LINT;
  bBuffer_Send  : ARRAY[0..1023] OF BYTE;
  bSendWatchDog : BOOL;
  mhMsgHeader   : MsgHeader;
  bSendMsgBlock : BOOL;
  pbCurPos_Send      : POINTER TO BYTE;
  bSendControlSystem : BOOL;
  bSendIoSystem      : BOOL;
  bSendDrives        : BOOL;
  SpsToTcp : SPSTOMMI;
  dwCrcTemp: DWORD;

  tnSendIoSystem: TON;
  tSendIoSystem: TIME := T#500MS;
  wSendIoSystem: WORD;
  wSendControlSystem: WORD;
  wSendMsgBlock: WORD;

  //ReadMsg
  l_b_ReadMsg_NewMsg : BOOL;
  l_b_ReadMsg_Body : BOOL;
  l_b_ReadMsg_Failure : BOOL;
END_VAR

TCP_Server();
END_FUNCTION_BLOCK

(* ---- TCPMain.prg.st ---- *)
(* METADATA
{
	"v3Meta": {
		"objectGuid": "bf44ddad-4c4e-44de-9f11-5004840b8d3d"
	}
}
*)
PROGRAM TCPMain
VAR_INPUT
  bpIOAnzeigeAktivieren : BOOL;
  l_fb_SortjetHMI : Hegla_Gateway_Komm_FB;
END_VAR
VAR
  bInit : BOOL := TRUE;
END_VAR

// MAIN PRG
IF bInit
THEN
  RegisterCallbacks();
  bInit := FALSE;
END_IF

l_fb_SortjetHMI();
END_PROGRAM
